*)
VAR_INPUT
	(* Variables *)
	bEnable								:BOOL;						(* Enable FB *)
	lrInSignal								:LREAL;						(* Input value to the block *)
	lrKp									:LREAL := 1;					(* Proportional gain of integrator *)
	tT1									:TIME := t#200ms;				(* Time constant  of integrator *)
	tTaskCycle							:TIME := t#2ms;				(* Cycle time *)
END_VAR
VAR_OUTPUT
	(* Variables *)
	lrOutSignal							:LREAL;						(* Output value the block state *)
END_VAR
VAR
	(* Variables *)
	bFirstTime							:BOOL;
	lrTimeRatio							:LREAL;

	lrLastSignal							:LREAL;						(* Last signal *)
END_VAR

IF NOT bEnable
THEN
	lrOutSignal := 0.0;
	bFirstTime := FALSE;
	RETURN;
END_IF


IF NOT bFirstTime
     OR tT1= t#0ms
     OR tT1 < (tTaskCycle + tTaskCycle)
THEN
	lrOutSignal := lrKp * lrInSignal;

	bFirstTime := TRUE;
ELSE
	lrTimeRatio := TIME_TO_LREAL(tTaskCycle) / TIME_TO_LREAL(tT1);

	lrOutSignal := (lrKp * lrInSignal * lrTimeRatio) + (lrLastSignal * (1 -  lrTimeRatio));
END_IF

lrLastSignal := lrOutSignal;

END_FUNCTION_BLOCK

// ---- POUs/Tc2 Objects/Engineering/Position offset/F_PosOffset.TcPOU
FUNCTION F_PosOffset : LREAL
(*

The function used to calculate position offset in range.

Constructor: 		Patryk Panylo
Company:		E. Riexinger GmbH
Date:			01.04.2015
Version:			1.00

Date:			Revision:		Who:				Comment
dd.mm.yyyy		x.xx			Initials			comment

*)
VAR_INPUT
	(* Input variables / Eingang Variablen *)
	bEnable							:BOOL;						(* Function enable *)
	lrCurrentPosHorizontal				:LREAL;						(* Current position of horizontal axis *)
	lrPosOffsetHorizontal				:LREAL;						(* Position offset of horizontal axis*)
	lrPosOffsetVertical					:LREAL;						(* Position offset of horizontal axis*)
	lrRangeOffset						:LREAL;						(* Range offset *)
END_VAR
VAR
	(* Variables *)

END_VAR

IF NOT bEnable
THEN
	F_PosOffset := 0.0;

	RETURN;
END_IF

IF  lrRangeOffset > 0.0
     AND lrCurrentPosHorizontal >= lrPosOffsetHorizontal - ABS(lrRangeOffset * 0.5)
     AND lrCurrentPosHorizontal <= lrPosOffsetHorizontal + ABS(lrRangeOffset * 0.5)
THEN
	F_PosOffset := lrPosOffsetVertical;
ELSE
	F_PosOffset := 0.0;
END_IF

END_FUNCTION

// ---- POUs/Tc2 Objects/Engineering/Position/F_ModuloDistance.TcPOU
FUNCTION F_ModuloDistance : DINT
(*
Function for calculate modulo distance.

Constructor: 	Patryk Panylo
Company:		E. Riexinger GmbH
Date:			20.01.2014
Version:		1.00

Date:			Revision:		Who:				Comment
dd.mm.yyyy		x.xx			Initials			comment

*)

VAR_INPUT
	dwCurrentValue			:DWORD;
	dwOldValue				:DWORD;
	dwModuloValue			:DWORD;
END_VAR
VAR
	dwPosDistance			:DWORD;

END_VAR


F_ModuloDistance := DWORD_TO_DINT(dwCurrentValue - dwOldValue);

IF dwModuloValue <> 0
THEN
	dwPosDistance := F_ModDW(dwCurrentValue - dwOldValue, dwModuloValue);
	
	F_ModuloDistance := DWORD_TO_DINT(dwPosDistance);
	
	IF dwPosDistance > (dwModuloValue / 2) 
	THEN
		F_ModuloDistance := -DWORD_TO_DINT(dwModuloValue - dwPosDistance);
	END_IF
	
END_IF

END_FUNCTION

// ---- POUs/Tc2 Objects/Mathematical/F_ModDW.TcPOU
FUNCTION F_ModDW : DWORD
(*
Modulo function for double word numbers (dividend mod divisor).

Constructor: 		Patryk Panylo
Company:		E. Riexinger GmbH
Date:			20.01.2014
Version:			1.00

Date:			Revision:		Who:				Comment
dd.mm.yyyy		x.xx			Initials			comment

*)
VAR_INPUT
	dwDividend						:DWORD;
	dwDivisor						:DWORD;
END_VAR
VAR
END_VAR


F_MODDW := dwDivisor;

IF dwDivisor <> 0 
THEN
	F_MODDW := dwDividend MOD dwDivisor;
END_IF;

END_FUNCTION

// ---- POUs/Tc2 Objects/Engineering/Trajectory model/FB_ExtContour.TcPOU
FUNCTION_BLOCK FB_ExtContour
(*

The function block used to generate move external contour.

Constructor: 		Patryk Panylo
Company:		E. Riexinger GmbH
Date:			01.04.2015
Version:			1.00

Date:			Revision:		Who:				Comment
dd.mm.yyyy		x.xx			Initials			comment

*)
VAR_INPUT
	(* Input variables / Eingang Variablen *)
	bEnable							:BOOL;						(* Function block enable *)
	bStart							:BOOL;
	bStop							:BOOL;
	etContourType					:ET_ContourType;				(* Contour type *)
	lrActPosZ						:LREAL;						(* Current position of axis z *)
	lrActAngle 						:LREAL; 						(* Current angle *)
	lrStartMaxPosZ					:LREAL;						(* Contour start maximal position of axis z *)
	lrEndMinPosZ					:LREAL;						(* Contour end minimal position of axis z *)
	lrSafetyDistance					:LREAL;						(* Safety distance *)
	lrTargetPosY						:LREAL;						(* Target position of axis y *)
END_VAR
VAR_OUTPUT
	(* Output variables / Ausgang Variablen *)
	lrNewPos						:LREAL;						(* New position [mm] *)
	bEnabled  						:BOOL;						(* Calculate positon is enabled *)
	lrActVelo							:LREAL;
	lrActPosN1						:LREAL;
END_VAR
VAR_IN_OUT
	lrSetPosY						:LREAL;						(* Set position of axis y *)
END_VAR
VAR
	(* Instances / Instanzen *)

	(* Enumerator  *)

	(* General flags / Allgemeine Variablen *)
	lrContourPos						:LREAL;
	bFirstTime						:BOOL;


END_VAR
VAR CONSTANT

END_VAR

IF NOT bEnable
THEN
	bEnabled := bStart;

	bFirstTime := FALSE;
	RETURN;
END_IF

IF NOT bFirstTime
THEN
	bEnabled := FALSE;

	bFirstTime := TRUE;
END_IF


IF bStop
THEN
	bEnabled := FALSE;

ELSIF bStart
THEN
	lrContourPos := F_CalcContour(
		etContourType := etContourType,
		lrActPos := lrActPosZ,
		lrActAngle := lrActAngle,
		(*lrActVelo := Axis.stNcToPlc.stCommandPositioning.dnActVelocity,*)
		lrVerticalOffset := 0.0,  (*37.0,*) (* Offset Sägeband Unterkante zu Störkontur BF-Kopf *)
		lrStartMaxPos := lrStartMaxPosZ,
		lrEndMinPos := lrEndMinPosZ,
		lrSafetyDistance := lrSafetyDistance,
		lrTableHeight := SEL(lrStartMaxPosZ>450, 700.0, 200.0), (* ab welcher Höhe Tischbreite aktiv ist *)
		lrTableWidth := 700.0, (* Tischbreite Auflage Rohr *)
		lrActVeloExt := lrActVelo
	);


	lrSetPosY := lrTargetPosY + lrContourPos;

	bEnabled := TRUE;

END_IF



lrActVelo := (*lrActVelo *0.9 + 0.1 *)(lrActPosZ - lrActPosN1);
lrActPosN1:= lrActPosZ;

END_FUNCTION_BLOCK

// ---- POUs/Tc2 Objects/Engineering/Trajectory model/F_CalcContour.TcPOU
FUNCTION F_CalcContour : LREAL
(*

The function used to calculate a contour of half circle dependent on angle of inclination axis and radius circle
Calculated position of axis is on output mapped.

Constructor: 		Patryk Panylo
Company:		E. Riexinger GmbH
Date:			01.04.2015
Version:			1.00

Date:			Revision:		Who:				Comment
dd.mm.yyyy		x.xx				Initials				comment
19.11.2015		1.01				ES					ET_ContourType_eEllipse
23.11.2015		1.02				ES					Square: also depending on angle(lrActAngle),
													lrVerticalOffset: guiding collision point is higher than act. position.

*)
VAR_INPUT
	(* Input variables / Eingang Variablen *)
	etContourType					:ET_ContourType;
	lrActPos							:LREAL;						(* Current position of axis *)
	lrActAngle						:LREAL;						(* Current angle, cutting angle *)
	(*lrActVelo							:LREAL;						(* Current speed of axis *)*)
	lrVerticalOffset					:LREAL;						(* vertical offset collision contour *)
	lrStartMaxPos						:LREAL;						(* Contour start maximal position *)
	lrEndMinPos						:LREAL;						(* Contour end minimal position  *)
	lrSafetyDistance					:LREAL;						(* Safety distance *)
	lrTableHeight						:LREAL;						(* Table height, if need guidings go to table width *)
	lrTableWidth						:LREAL;						(* table width *)
	lrActVeloExt						:LREAL;						(* Current velo of axis *)
END_VAR
VAR
	(* Variables *)
	lrActPosCache					:LREAL;						(* intern position of axis *)
	lrRadius							:LREAL;						(* Radius *)
	lrMiddlePos						:LREAL;						(* Middle position *)
	lrAlfa							:LREAL;						(* Angle of inclination *)
	lrDelta							:LREAL;						(* Distance z = f(x)*)
	lrCosAlfa							:LREAL;						(* Cosine of alfa *)
	lrAngleFactor						:LREAL;						(* Sawbow angle factor, ellipse *)
	lrStartMaxPosCache 				:LREAL;
	lrEndMinPosCache 				:LREAL;

END_VAR

lrStartMaxPosCache := lrStartMaxPos + ABS(lrSafetyDistance) + 50.0;
lrEndMinPosCache := lrEndMinPos - ABS(lrSafetyDistance) + 50.0;

lrActPosCache := lrActPos - lrVerticalOffset;

CASE etContourType OF

	ET_ContourType_eNone:
		F_CalcContour := lrActPosCache;

	ET_ContourType_eCircle, ET_ContourType_eEllipse:
		lrRadius := ABS(lrStartMaxPosCache - lrEndMinPos) / 2;
		lrMiddlePos := lrEndMinPosCache + lrRadius;										(* Middle position *)

		IF (lrActPosCache <= lrStartMaxPosCache)
		     AND (lrActPosCache >= lrEndMinPosCache)
		     AND lrRadius > 0.0
		THEN
			lrAlfa := ASIN(ABS(lrActPosCache - lrMiddlePos) /  lrRadius);				(* Angle of inclination *)
			lrCosAlfa := COS(lrAlfa);												(* Cosine of alfa *)
			lrDelta := lrCosAlfa * lrRadius;								(* Distance z = f(x)*)

			F_CalcContour := lrDelta;

		ELSE
			F_CalcContour := 0.0;
		END_IF

		IF lrActPos <= lrTableHeight
			OR lrActPos < lrMiddlePos
		THEN
			F_CalcContour := MAX(F_CalcContour, lrTableWidth / 2 + lrSafetyDistance);
		END_IF

		IF ((lrActVeloExt>0.0)
			AND (lrActPosCache < lrMiddlePos))
			OR ((lrActVeloExt=0.0)
			AND lrActPos < lrTableHeight)
		THEN
			F_CalcContour := MAX(lrRadius, lrTableWidth / 2 + lrSafetyDistance);
		END_IF

		IF etContourType = ET_ContourType_eEllipse
		THEN
			lrAngleFactor := 1 /  COS( MIN(ABS(lrActAngle), 89.9) / 180.0*PI);
			F_CalcContour := F_CalcContour * lrAngleFactor;
		END_IF

	ET_ContourType_eSquare:
		lrRadius := ABS(lrStartMaxPosCache - lrEndMinPos) / 2;
		lrMiddlePos := lrEndMinPosCache + lrRadius;										(* Middle position *)

		IF (lrActPosCache <= lrStartMaxPosCache)
		     AND (lrActPosCache >= lrEndMinPosCache)
		     AND lrRadius > 0.0
		THEN
			lrDelta := lrRadius;													(* Distance z = f(x)*)

			F_CalcContour := lrDelta;

		ELSE
			F_CalcContour := 0.0;
		END_IF

		IF lrActPos <= lrTableHeight
		THEN
			F_CalcContour := MAX(F_CalcContour, lrTableWidth / 2 + lrSafetyDistance / 2);
		END_IF

		lrAngleFactor := 1 /  COS( MIN(ABS(lrActAngle), 89.9) / 180.0*PI);
		F_CalcContour := F_CalcContour * lrAngleFactor;

ELSE
	F_CalcContour := 0.0;

END_CASE;

END_FUNCTION

// ---- POUs/Tc2 Objects/Engineering/Trajectory model/FB_ExtTraj.TcPOU
FUNCTION_BLOCK FB_ExtTraj
(*

The function block used to generate move external trajectory.

Constructor: 		Patryk Panylo
Company:		E. Riexinger GmbH
Date:			01.04.2015
Version:			1.00

Date:			Revision:		Who:				Comment
dd.mm.yyyy		x.xx			Initials			comment

*)
VAR_INPUT
	(* Input variables / Eingang Variablen *)
	bEnable							:BOOL;						(* Function block enable *)
	bStart							:BOOL;						(* Execute start an external trajectory with rising edge *)
	bStop							:BOOL;						(* Execute stop an external trajectory with rising edge *)
	lrStartPosHorizontal				:LREAL;						(* Start position of horizontal axis [mm] *)
	lrStartPosVertical					:LREAL;						(* Start position of vertical axis [mm] *)
	lrRadius							:LREAL;						(* Radius of circle [mm] *)
	unPosWindow					:UINT := 2;					(* Position window [mm] *)
	bTakeHorMovePara				:BOOL;						(* Take move parameters from 1- horizontal axis, 0 - vertical axis *)
END_VAR
VAR_OUTPUT
	(* Output variables / Ausgang Variablen *)
	lrNewPos						:LREAL;						(* New position [mm] *)
	lrNewVelo						:LREAL;						(* New velocity [mm/s] *)
	lrNewAcc						:LREAL;						(* New acceleration [mm/s^2] *)
	bEnabled  						:BOOL;						(* Calculate positon is enabled *)
	bDone							:BOOL;						(* Command done *)
	bBusy							:BOOL;						(* Command busy *)
	bError							:BOOL;						(* Command error  *)
	udnErrorNo						:UDINT;						(* Error number *)
	sErrorMsg						:STRING; 					(* Error message *)
END_VAR
VAR_IN_OUT
	AxisHorizontal					:AXIS_REF;					(* The AXIS_REF data type  is an interface between the PLC and the NC and contains axis information *)
	AxisVertical						:AXIS_REF;					(* The AXIS_REF data type  is an interface between the PLC and the NC and contains axis information *)
END_VAR
VAR
	(* Instances / Instanzen *)

	(* Enumerator  *)
	etCalcExtTrajState					:ET_CalcExtTrajState;								(* Current state *)

	(* General flags / Allgemeine Variablen *)
	lrExtStartPosHorizontal				:LREAL;
	lrExtStartPosVertical				:LREAL;
	lrExtRadius						:LREAL;

	bFirstTime						:BOOL;
END_VAR
VAR CONSTANT

END_VAR

IF NOT bEnable
THEN
	lrNewPos := SEL(bTakeHorMovePara, AxisVertical.NcToPlc.SetPos, AxisHorizontal.NcToPlc.SetPos);
	lrNewVelo := SEL(bTakeHorMovePara, AxisVertical.NcToPlc.SetVelo, AxisHorizontal.NcToPlc.SetVelo);
	lrNewAcc := SEL(bTakeHorMovePara, AxisVertical.NcToPlc.SetAcc, AxisHorizontal.NcToPlc.SetAcc);

	bDone := FALSE;					(* Command done *)
	bBusy := FALSE;					(* Command busy *)
	bError := FALSE;					(* Command error  *)
	udnErrorNo := 0;					(* Error number *)
	sErrorMsg := ''; 					(* Error message *)

	bEnabled := FALSE;

	bFirstTime := FALSE;
	RETURN;
END_IF

IF NOT bFirstTime
THEN
	bEnabled := FALSE;

	etCalcExtTrajState := ET_CalcExtTrajState_eWaitExecute;

	bFirstTime := TRUE;
END_IF

CASE etCalcExtTrajState
OF
	ET_CalcExtTrajState_eWaitExecute:
		IF bStop
		THEN
			bEnabled := FALSE;

			bDone := FALSE;						(* Command done *)
			bBusy := TRUE;						(* Command busy *)
			bError := FALSE;						(* Command error  *)
			udnErrorNo := 0;						(* Error number *)
			sErrorMsg := ''; 						(* Error message *)

			etCalcExtTrajState := ET_CalcExtTrajState_eDone;

		ELSIF bStart
		THEN
			bDone := FALSE;						(* Command done *)
			bBusy := TRUE;						(* Command busy *)
			bError := FALSE;						(* Command error  *)
			udnErrorNo := 0;						(* Error number *)
			sErrorMsg := ''; 						(* Error message *)

			etCalcExtTrajState := ET_CalcExtTrajState_eCalcTrajPos;

		END_IF

	ET_CalcExtTrajState_eCalcTrajPos:
		bEnabled := TRUE;

		lrExtStartPosHorizontal := lrStartPosHorizontal;
		lrExtStartPosVertical := lrStartPosVertical;
		lrExtRadius := lrRadius;

		etCalcExtTrajState := ET_CalcExtTrajState_eDone;

	ET_CalcExtTrajState_eError:
		bBusy := FALSE;						(* Command busy *)
		bError := TRUE;						(* Command error  *)

		etCalcExtTrajState := ET_CalcExtTrajState_eNoExecute;

	ET_CalcExtTrajState_eDone:
		bDone := TRUE;						(* Command done *)
		bBusy := FALSE;						(* Command busy *)

		etCalcExtTrajState := ET_CalcExtTrajState_eNoExecute;

	ET_CalcExtTrajState_eNoExecute:
		IF NOT bStart
		     AND NOT bStop
		THEN
			(* Reset outputs *)
			bDone := FALSE;						(* Command done *)
			bBusy := FALSE;						(* Command busy *)
			bError := FALSE;						(* Command error  *)

			etCalcExtTrajState := ET_CalcExtTrajState_eWaitExecute;
		END_IF
END_CASE

(* The function is used to calculate a trajectory of vertical position. *)
IF bEnabled
THEN
	lrNewPos := F_CalcTrajPos(
		lrStartPosHorizontal := lrExtStartPosHorizontal,
		lrStartPosVertical := lrExtStartPosVertical,
		lrCurrentPosHorizontal := AxisHorizontal.NcToPlc.SetPos,
		lrCurrentPosVertical := AxisVertical.NcToPlc.SetPos,
		lrRadius := lrExtRadius
	);

	lrNewVelo := AxisHorizontal.NcToPlc.SetVelo;
	lrNewAcc := AxisHorizontal.NcToPlc.SetAcc;

	(* ABS(lrNewPos - AxisVertical.NcToPlc.SetPos) > UINT_TO_LREAL(unPosWindow)
	THEN
		bError := TRUE;								(* Command error  *)
		udnErrorNo :=  1;								(* Error number *)
		sErrorMsg := ''; 								(* Error message *)
	END_IF*)
ELSE
	lrNewPos := SEL(bTakeHorMovePara, AxisVertical.NcToPlc.SetPos, AxisHorizontal.NcToPlc.SetPos);
	lrNewVelo := SEL(bTakeHorMovePara, AxisVertical.NcToPlc.SetVelo, AxisHorizontal.NcToPlc.SetVelo);
	lrNewAcc := SEL(bTakeHorMovePara, AxisVertical.NcToPlc.SetAcc, AxisHorizontal.NcToPlc.SetAcc);

	bError := FALSE;								(* Command error  *)
	udnErrorNo :=  0;								(* Error number *)
	sErrorMsg := ''; 								(* Error message *)
END_IF

END_FUNCTION_BLOCK

// ---- POUs/Tc2 Objects/Engineering/Trajectory model/F_CalcTrajPos.TcPOU
FUNCTION F_CalcTrajPos : LREAL
(*

The function used to calculate a trajectory of half circle dependent on angle of inclination axis and radius circle
Calculated position of axis is on output mapped.

Constructor: 		Patryk Panylo
Company:		E. Riexinger GmbH
Date:			01.04.2015
Version:			1.00

Date:			Revision:		Who:				Comment
dd.mm.yyyy		x.xx			Initials			comment

*)
VAR_INPUT
	(* Input variables / Eingang Variablen *)
	lrStartPosHorizontal				:LREAL;						(* Start position of horizontal axis *)
	lrStartPosVertical					:LREAL;						(* Start position of vertical axis *)
	lrCurrentPosHorizontal				:LREAL;						(* Current position of horizontal axis *)
	lrCurrentPosVertical				:LREAL;						(* Current position of vertical axis *)
	lrRadius							:LREAL;						(* Radius of circle *)
END_VAR
VAR
	(* Variables *)
	lrAlfa							:LREAL;						(* Angle of inclination *)
	lrDelta							:LREAL;						(* Distance z = f(x)*)
	lrCosAlfa							:LREAL;						(* Cosine of alfa *)
END_VAR

IF lrRadius > 0.0
THEN
	IF ABS(lrCurrentPosHorizontal - lrStartPosHorizontal) / lrRadius <= 1.0
	THEN
		lrAlfa := ASIN(ABS(lrCurrentPosHorizontal - lrStartPosHorizontal) / lrRadius);					(* Angle of inclination *)
		lrCosAlfa := COS(lrAlfa);																(* Cosine of alfa *)
		lrDelta := lrRadius - (lrCosAlfa * lrRadius);											(* Distance z = f(x)*)

		F_CalcTrajPos := lrCurrentPosVertical - lrDelta;
	ELSE
		F_CalcTrajPos := lrCurrentPosVertical;
	END_IF
ELSE
	F_CalcTrajPos := lrCurrentPosVertical;
END_IF

END_FUNCTION

// ---- POUs/Tc2 Objects/ExternalHardware/Gefran/FB_GFX4IRCtrlZone.TcPOU
FUNCTION_BLOCK FB_GFX4IRCtrlZone
(*

The function block used to control Gerfan GFX4IR zone.

Constructor: 		Patryk Panylo
Company:		E. Riexinger GmbH
Date:			12.07.2016
Version:			1.00

Date:			Revision:		Who:				Comment
13.12.2017		1.01				PPA					Control with temperatur feedback

*)
VAR_INPUT
	(* Input variables / Eingang Variablen *)
	bEnable							:BOOL;						(* Function block enable *)
	bReset							:BOOL;						(* Controller reset *)
	bHandStart						:BOOL;						(* Execute start an external trajectory with rising edge *)
	bHandStop						:BOOL;						(* Execute stop an external trajectory with rising edge *)
	bAutoStart						:BOOL;						(* Execute start an external trajectory with rising edge *)
	bAutoStop						:BOOL;						(* Execute stop an external trajectory with rising edge *)
	bStartRelease					:BOOL;						(* Start release *)
	bCtrlInterrupt						:BOOL;						(* Control interrupt *)
	lrSetpoint						:LREAL;						(* Setpoint *)
	bCtrlManAuto						:BOOL;						(* Auto := FALSE, Man := TRUE *)
	bEnAutoCtrlOff					:BOOL := TRUE;				(* Auto off enable*)
	tControllerOff						:TIME := t#90s;				(* Time to switch controller off *)
	tControllerOn						:TIME := t#90s;				(* Time to switch controller on *)
	lrTempMin						:LREAL;						(* Minimal temperature *)
	lrTempMax						:LREAL;						(* Maximal temperature *)
	lrTempLimitMin					:LREAL;						(* Minimal temperature limit *)
	lrTempLimitMax					:LREAL;						(* Maximal temperature limit *)
END_VAR
VAR_OUTPUT
	(* Output variables / Ausgang Variablen *)
	unCurrentValue					:UINT;						(* Current value *)
	bEnabled  						:BOOL;						(* Zone enabled *)
	bDamaged						:BOOL;						(* Zone damaged *)
	bDone							:BOOL;						(* Command done *)
	bBusy							:BOOL;						(* Command busy *)
	bError							:BOOL;						(* Command error  *)
	udnErrorNo						:UDINT;						(* Error number *)
	sErrorMsg						:STRING; 					(* Error message *)
END_VAR
VAR_IN_OUT
	(* Input Output variables / Ausgang Variablen *)
	CtrlGFX4IRTOPLC					:ST_GFX4IRTOPLC;			(* The ST_GFX4IRTOPLC data type  is an interface between the PLC and the GFX4IR and contains controller information *)
	CtrlPLCTOGFX4IR					:ST_PLCTOGFX4IR;			(* The ST_PLCTOGFX4IR data type  is an interface between the PLC and the GFX4IR and contains controller information *)
END_VAR
VAR
	(* Enummerations *)
	etGFX4IRStates					:ET_GFX4IR := ET_GFX4IRState_eWaitExecute;			(* Current state *)

	(* Variables *)
	nWatchdog						:INT;
	bControllerOn						:BOOL;

	bFirstTime						:BOOL;

	(* References *)

	(* Interfaces *)

	(* Instances *)
	fbControllerOff					:FB_SignalHandlingDelay;
	fbControllerOn					:FB_SignalHandlingDelay;
	fbScalingSP						:FB_Scaling;

	rtAutoStart						:R_TRIG;
	rtAutoStop						:R_TRIG;
	rtHandStart						:R_TRIG;
	rtHandStop						:R_TRIG;
END_VAR
VAR CONSTANT

END_VAR


IF NOT bFirstTime
THEN
	bControllerOn := TRUE;

	nWatchdog := 0;
	bDone := FALSE;						(* Command done *)
	bBusy := FALSE;						(* Command busy *)
	bError := FALSE;						(* Command error  *)

	etGFX4IRStates := ET_GFX4IRState_eWaitExecute;

	bFirstTime := TRUE;
END_IF

(* Scaling set point *)
fbScalingSP(
	bEnable := TRUE,
	lrInput := lrSetpoint,
	lrXLowLimit := lrTempMin,
	lrXUpperLimit := lrTempMax,
	lrYLowLimit := lrTempLimitMin,
	lrYUpperLimit := lrTempLimitMax,
	usiPrecision := 2
);

CtrlPLCTOGFX4IR.wControllerStatus.4 := bCtrlManAuto;			(* Auto := FALSE, Man := TRUE *)

IF bCtrlManAuto										(* Auto := FALSE, Man := TRUE *)
THEN
	bEnabled := CtrlGFX4IRTOPLC.nOutputPower > 0
			       AND (CtrlGFX4IRTOPLC.nOutputPower = LREAL_TO_INT(lrSetpoint  * 10.0));
			       (*AND CtrlGFX4IRTOPLC.wControllerStatus.5					(* Ctrl enabled  *)
			          AND NOT CtrlGFX4IRTOPLC.wControllerStatus.0;			(* Alarm  *)*)
ELSE
	bEnabled := CtrlGFX4IRTOPLC.nOutputPower > 0;
			       (*AND (CtrlGFX4IRTOPLC.nProcessVariable >= LREAL_TO_INT(fbScalingSP.lrOutputPV));*)
			       (*AND CtrlGFX4IRTOPLC.wControllerStatus.5					(* Ctrl enabled  *)
			          AND NOT CtrlGFX4IRTOPLC.wControllerStatus.0;			(* Alarm  *)*)
END_IF

bDamaged := CtrlGFX4IRTOPLC.wControllerStatus.12;
unCurrentValue := CtrlGFX4IRTOPLC.nOutputPower / 10;

fbControllerOff(
	bEnable := TRUE,
	bIn := bEnAutoCtrlOff
		  AND bEnabled,
	tDelay := tControllerOff
);

fbControllerOn(
	bEnable := TRUE,
	bIn := NOT bEnabled					(* Ctrl disabled *)
		  AND NOT bControllerOn,
	tDelay := tControllerOn
);

(*
IF bHandStop
    OR bCtrlInterrupt
THEN
	CtrlPLCTOGFX4IR.wControllerStatus.3 := TRUE;			(* Ctrl ON = FALSE, OFF = TRUE *)
	CtrlPLCTOGFX4IR.nLocalSetPoint := 0;
	CtrlPLCTOGFX4IR.nManualOutput := 0;
ELSIF bHandStart
THEN
	CtrlPLCTOGFX4IR.wControllerStatus.3 := FALSE;			(* Ctrl ON = FALSE, OFF = TRUE *)
	CtrlPLCTOGFX4IR.nManualOutput := LREAL_TO_INT(lrSetpoint  * 10);
END_IF

RETURN;
*)

IF bCtrlInterrupt
     OR fbControllerOff.bOut
THEN
	bControllerOn := FALSE;

	CtrlPLCTOGFX4IR.wControllerStatus.3 := TRUE;			(* Ctrl ON = FALSE, OFF = TRUE *)
	CtrlPLCTOGFX4IR.nLocalSetPoint := 0;
	CtrlPLCTOGFX4IR.nManualOutput := 0;

	nWatchdog := 0;
	bDone := FALSE;						(* Command done *)
	bBusy := FALSE;						(* Command busy *)
	bError := FALSE;						(* Command error  *)

	etGFX4IRStates := ET_GFX4IRState_eWaitExecute;

ELSIF fbControllerOn.bOut
THEN
	bControllerOn := TRUE;
END_IF

IF bReset
     AND bError
THEN
	(* Reset outputs *)
	nWatchdog := 0;
	bDone := FALSE;						(* Command done *)
	bBusy := FALSE;						(* Command busy *)
	bError := FALSE;						(* Command error  *)

	etGFX4IRStates := ET_GFX4IRState_eWaitExecute;
ELSE
	(*IF bEnable
	     AND CtrlGFX4IRTOPLC.wControllerStatus.8					(* Ctrl error *)
	THEN
		bError := TRUE;									(* Command error  *)

		etGFX4IRStates := ET_GFX4IRState_eError;             		(* Next step *)
	END_IF*);
END_IF

rtHandStart(CLK := bHandStart);
rtHandStop(CLK := bHandStop);
rtAutoStart(CLK := bAutoStart AND bStartRelease AND bControllerOn);
rtAutoStop(CLK := bAutoStop);

IF rtHandStart.Q OR rtHandStop.Q
     OR rtAutoStart.Q OR rtAutoStop.Q
THEN
	nWatchdog := 0;
	bDone := FALSE;						(* Command done *)
	bBusy := FALSE;						(* Command busy *)
	bError := FALSE;						(* Command error  *)

	etGFX4IRStates := ET_GFX4IRState_eWaitExecute;
END_IF

CASE etGFX4IRStates
OF
	ET_GFX4IRState_eWaitExecute:
		IF NOT bEnable
		THEN
			bDone := TRUE;						(* Command done *)
			bBusy := TRUE;						(* Command busy *)
			bError := FALSE;						(* Command error  *)
			bEnabled  := bAutoStart AND NOT bAutoStop; 				(* Controller enabled *)

			etGFX4IRStates := ET_GFX4IRState_eWaitExecute;

		ELSIF NOT bCtrlInterrupt
			    AND NOT fbControllerOff.bOut
		THEN
			IF bAutoStop
			     OR bHandStop
			THEN
				nWatchdog := 0;

				bDone := FALSE;						(* Command done *)
				bBusy := TRUE;						(* Command busy *)
				bError := FALSE;						(* Command error  *)
				udnErrorNo := 0;						(* Error number *)
				sErrorMsg := ''; 						(* Error message *)

				etGFX4IRStates := ET_GFX4IRState_eCtrlOff;

			ELSIF rtAutoStart.Q
				    OR (rtHandStart.Q
					    AND bStartRelease
					    AND bControllerOn)
			THEN
				nWatchdog := 0;

				bDone := FALSE;						(* Command done *)
				bBusy := TRUE;						(* Command busy *)
				bError := FALSE;						(* Command error  *)
				udnErrorNo := 0;						(* Error number *)
				sErrorMsg := ''; 						(* Error message *)

				etGFX4IRStates := ET_GFX4IRState_eCtrlOn;

			END_IF
		END_IF

	ET_GFX4IRState_eCtrlOn:
		nWatchdog := nWatchdog + 1;

		CtrlPLCTOGFX4IR.wControllerStatus.3 := FALSE;			(* Ctrl ON = FALSE, OFF = TRUE *)

		IF bCtrlManAuto										(* Auto := FALSE, Man := TRUE *)
		THEN
			CtrlPLCTOGFX4IR.nManualOutput := LREAL_TO_UINT(lrSetpoint  * 10.0);
		ELSE
			CtrlPLCTOGFX4IR.nLocalSetPoint := LREAL_TO_INT(fbScalingSP.lrOutputPV);
		END_IF

		IF bEnabled											(* Ctrl enabled *)
		THEN
			nWatchdog := 0;
			etGFX4IRStates := ET_GFX4IRState_eDone;

		ELSIF nWatchdog > 5000
		THEN
			CtrlPLCTOGFX4IR.wControllerStatus.3 := TRUE;			(* Ctrl ON = FALSE, OFF = TRUE *)

			etGFX4IRStates := ET_GFX4IRState_eError;            		 (* Next step *)
		END_IF

	ET_GFX4IRState_eCtrlOff:
		nWatchdog := nWatchdog + 1;

		CtrlPLCTOGFX4IR.wControllerStatus.3 := TRUE;			(* Ctrl ON = FALSE, OFF = TRUE *)
		CtrlPLCTOGFX4IR.nLocalSetPoint := 0;
		CtrlPLCTOGFX4IR.nManualOutput := 0;

		IF NOT bEnabled
		THEN
			nWatchdog := 0;
			etGFX4IRStates := ET_GFX4IRState_eDone;

		ELSIF nWatchdog > 1000
		THEN
			CtrlPLCTOGFX4IR.wControllerStatus.3 := TRUE;			(* Ctrl ON = FALSE, OFF = TRUE *)
			CtrlPLCTOGFX4IR.nLocalSetPoint := 0;
			CtrlPLCTOGFX4IR.nManualOutput := 0;
			etGFX4IRStates := ET_GFX4IRState_eError;             		(* Next step *)
		END_IF

	ET_GFX4IRState_eDone:
		nWatchdog := 0;
		bDone := TRUE;						(* Command done *)
		bBusy := FALSE;						(* Command busy *)

		etGFX4IRStates := ET_GFX4IRState_eNoExecute;

	ET_GFX4IRState_eError:
		nWatchdog := 0;
		bBusy := FALSE;						(* Command busy *)
		bError := TRUE;						(* Command error  *)

		CtrlPLCTOGFX4IR.wControllerStatus.3 := TRUE;			(* Ctrl ON = FALSE, OFF = TRUE *)
		CtrlPLCTOGFX4IR.nLocalSetPoint := 0;
		CtrlPLCTOGFX4IR.nManualOutput := 0;

		etGFX4IRStates := ET_GFX4IRState_eNoExecute;

	ET_GFX4IRState_eNoExecute:
		IF NOT bHandStart
		     AND NOT bHandStop
		     AND NOT bAutoStart
		     AND NOT bAutoStop
		THEN
			(* Reset outputs *)
			nWatchdog := 0;
			bDone := FALSE;						(* Command done *)
			bBusy := FALSE;						(* Command busy *)
			bError := FALSE;						(* Command error  *)

			etGFX4IRStates := ET_GFX4IRState_eWaitExecute;
		END_IF
END_CASE

END_FUNCTION_BLOCK

// ---- POUs/Tc2 Objects/ExternalHardware/Gefran/FB_GFX4IRZones.TcPOU
FUNCTION_BLOCK FB_GFX4IRZones
(*

The function block used to control Gerfan GFX4IR Zones.

Constructor: 		Patryk Panylo
Company:		E. Riexinger GmbH
Date:			12.07.2016
Version:			1.00

Date:			Revision:		Who:				Comment
25.09.2017		1.01				PPA					Change check zone damaged

*)
VAR_INPUT
	(* Input variables / Eingang Variablen *)
	bEnable							:BOOL;													(* Function block enable *)
	arbZoneEn						:ARRAY[1..nZONES_MAX_NO] OF BOOL;						(* Zone enable *)
	bReset							:BOOL;													(* Reset *)
	arbHandStart						:ARRAY[1..nZONES_MAX_NO] OF BOOL;						(* Execute start GFX4IR controller with rising edge *)
	arbHandStop						:ARRAY[1..nZONES_MAX_NO] OF BOOL;						(* Execute stop GFX4IR controller with rising edge *)
	bAutoStart						:BOOL;													(* Execute start GFX4IR controller with rising edge *)
	bAutoStop						:BOOL;													(* Execute stop GFX4IR controller with rising edge *)
	bStartRelease					:BOOL;													(* Start release *)
	bCtrlInterrupt						:BOOL;													(* Control interrupt *)
	arlrSetpoint						:ARRAY[1..nZONES_MAX_NO] OF LREAL;					(* Setpoint *)
	bCtrlManAuto						:BOOL;													(* Auto := FALSE, Man := TRUE *)
	bEnAutoCtrlOff					:BOOL := TRUE;											(* Auto controller off enable*)
	bEnOneByOneOn					:BOOL := FALSE;											(* One by one switch on *)
	tDelayZoneOn					:TIME := t#100ms;											(* Delay time of zone one by one to switch on *)
	tControllerOff						:TIME := t#90s;											(* Time to switch controller off *)
	tControllerOn						:TIME := t#90s;											(* Time to switch controller on *)
	lrTempMin						:LREAL;													(* Minimal temperature *)
	lrTempMax						:LREAL;													(* Maximal temperature *)
	lrTempLimitMin					:LREAL;													(* Minimal temperature limit *)
	lrTempLimitMax					:LREAL;													(* Maximal temperature limit *)
END_VAR
VAR_OUTPUT
	(* Output variables / Ausgang Variablen *)
	arunCurrentValue					:ARRAY[1..nZONES_MAX_NO] OF UINT;						(* Current value *)
	bEnabled  						:BOOL;													(* Zone enabled *)
	bEnabledDelay					:BOOL;													(* Zone enabled delay *)
	arbZoneDamaged				:ARRAY[1..nZONES_MAX_NO] OF BOOL;
	bDone							:BOOL;						(* Command done *)
	bError							:BOOL;						(* Command error  *)
	udnErrorNo						:UDINT;						(* Error number *)
END_VAR
VAR_IN_OUT
	(* Input Output variables / Ausgang Variablen *)
	GFX4IR							:ST_GFX4IR_REF;				(* The ST_GFX4IR_REF data type  is an interface between the PLC and the GFX4IR and contains controller information *)
END_VAR
VAR
	(* Enummerations *)

	(* Variables *)
	nIdx								:INT;
	tEnabledDelay					:TIME := t#1s;					(* Enabled delay time *)


	bFirstTime						:BOOL;

	(* References *)

	(* Interfaces *)

	(* Instances *)
	arfbGFX4IRCtrlZone				:ARRAY[1..nZONES_MAX_NO] OF FB_GFX4IRCtrlZone;
	tonEnabledDelay					:TON;						(* Delay controller enabled status *)
	tonDelayZoneOn					:ARRAY[1..nZONES_MAX_NO] OF TON;						(* Delay zone one by one to switch on *)

END_VAR


IF NOT bEnable
THEN
	bDone := FALSE;					(* Command done *)
	bError := FALSE;					(* Command error  *)

	FOR nIdx := 1 TO nZONES_MAX_NO
	DO
		arfbGFX4IRCtrlZone[nIdx](
			bEnable := TRUE,
			bAutoStart := bAutoStart,
			bAutoStop := bAutoStop,
			bCtrlInterrupt := bCtrlInterrupt,
			lrTempMin := lrTempMin,
			lrTempMax := lrTempMax,
			lrTempLimitMin := lrTempLimitMin,
			lrTempLimitMax := lrTempLimitMax,
			CtrlGFX4IRTOPLC := GFX4IR.Gfx4IRToPlc[nIdx],
			CtrlPLCTOGFX4IR := GFX4IR.PlcToGfx4IR[nIdx],
			unCurrentValue => arunCurrentValue[nIdx]
		 );
	END_FOR

	bEnabled := FALSE;
	bEnabledDelay := FALSE;

	bFirstTime := FALSE;
	RETURN;
END_IF

IF NOT bFirstTime
THEN
	bDone := FALSE;					(* Command done *)
	bError := FALSE;					(* Command error  *)

	bEnabled := FALSE;
	bEnabledDelay := FALSE;

	bFirstTime := TRUE;
END_IF

bEnabled := TRUE;
bDone := TRUE;
bError := FALSE;

FOR nIdx := 1 TO nZONES_MAX_NO
DO
	(*
	IF bAutoStart
	THEN
		IF bEnOneByOneOn
		     AND tDelayZoneOn > t#0ms
		     AND nIdx > 1
		     AND NOT arfbGFX4IRController[nIdx].bEnabled
		THEN
			tonDelayZoneOn[nIdx](
				IN := arfbGFX4IRController[nIdx - 1].bEnabled,
				PT := tDelayZoneOn
			);
	
			IF tonDelayZoneOn[nIdx].Q
			THEN
				arfbGFX4IRController[nIdx].bStartRelease := bStartRelease;
			ELSE
				arfbGFX4IRController[nIdx].bStartRelease := FALSE;;
			END_IF
		ELSE
			tonDelayZoneOn[nIdx](IN := FALSE);
			arfbGFX4IRController[nIdx].bStartRelease := bStartRelease;
		END_IF
	ELSE
		tonDelayZoneOn[nIdx](IN := FALSE);
		arfbGFX4IRController[nIdx].bStartRelease := bStartRelease;
	END_IF
	*)

	arfbGFX4IRCtrlZone[nIdx].bStartRelease := bStartRelease;

	arfbGFX4IRCtrlZone[nIdx](
		bEnable := arbZoneEn[nIdx],
		bReset := bReset,
		bHandStart := arbHandStart[nIdx],
		bHandStop := arbHandStop[nIdx],
		bAutoStart := bAutoStart,
		bAutoStop := bAutoStop,
		bCtrlInterrupt := bCtrlInterrupt,
		lrSetpoint := arlrSetpoint[nIdx],
		bCtrlManAuto := bCtrlManAuto,
		bEnAutoCtrlOff := bEnAutoCtrlOff,
		tControllerOff := tControllerOff,
		tControllerOn := tControllerOn,
		lrTempMin := lrTempMin,
		lrTempMax := lrTempMax,
		lrTempLimitMin := lrTempLimitMin,
		lrTempLimitMax := lrTempLimitMax,
		CtrlGFX4IRTOPLC := GFX4IR.Gfx4IRToPlc[nIdx],
		CtrlPLCTOGFX4IR := GFX4IR.PlcToGfx4IR[nIdx],
		unCurrentValue => arunCurrentValue[nIdx],
		bDamaged => arbZoneDamaged[nIdx]
	 );

	bEnabled := bEnabled AND arfbGFX4IRCtrlZone[nIdx].bEnabled;
	bDone := bDone AND arfbGFX4IRCtrlZone[nIdx].bDone;
	bError := bError OR arfbGFX4IRCtrlZone[nIdx].bError;

END_FOR

tonEnabledDelay(
	IN := bEnabled,
	PT := tEnabledDelay,
	Q => bEnabledDelay
);

END_FUNCTION_BLOCK

// ---- POUs/Tc2 Objects/ExternalHardware/Gefran/FB_GFX4IR_REF.TcPOU
FUNCTION_BLOCK FB_GFX4IR_REF
VAR_INPUT
	Gfx4IRToPlc			AT %I*:ARRAY[1..4] OF ST_GFX4IRTOPLC;
END_VAR
VAR_OUTPUT
	PlcToGfx4IR			AT %Q*:ARRAY[1..4] OF ST_PLCTOGFX4IR;
END_VAR
VAR
END_VAR

;

END_FUNCTION_BLOCK

// ---- POUs/Tc2 Objects/ExternalHardware/Gefran/F_ChkAllZonesNotEnabled.TcPOU
FUNCTION F_ChkAllZonesNotEnabled : BOOL
(*

The function used to detect if all controller are enabled.

Constructor: 		Patryk Panylo
Company:		E. Riexinger GmbH
Date:			23.04.2015
Version:			1.00

Date:			Revision:		Who:				Comment
dd.mm.yyyy		x.xx			Initials			comment

*)
VAR_INPUT
	(* Input variables / Eingang Variablen *)
	bEnable						:BOOL;						(* Signal FB enable *)
	GFX4IR1						:ST_GFX4IR_REF;				(* The ST_GFX4IRTOPLC data type  is an interface between the PLC and the GFX4IR and contains controller information *)
	GFX4IR2						:ST_GFX4IR_REF;				(* The ST_GFX4IRTOPLC data type  is an interface between the PLC and the GFX4IR and contains controller information *)
	GFX4IR3						:ST_GFX4IR_REF;				(* The ST_GFX4IRTOPLC data type  is an interface between the PLC and the GFX4IR and contains controller information *)
	GFX4IR4						:ST_GFX4IR_REF;				(* The ST_GFX4IRTOPLC data type  is an interface between the PLC and the GFX4IR and contains controller information *)
END_VAR
VAR
	(* Enummerations *)

	(* Variables *)

	(* References *)

	(* Interfaces *)

	(* Instances *)

END_VAR


IF NOT bEnable							(* Signal FB enable *)
THEN
	F_ChkAllZonesNotEnabled := FALSE;

	RETURN;
END_IF

F_ChkAllZonesNotEnabled := GFX4IR1.Gfx4IRToPlc[1].nProcessVariable = 0
						   AND GFX4IR1.Gfx4IRToPlc[2].nProcessVariable = 0
						   AND GFX4IR1.Gfx4IRToPlc[3].nProcessVariable = 0
						   AND GFX4IR1.Gfx4IRToPlc[4].nProcessVariable = 0
						   AND GFX4IR2.Gfx4IRToPlc[1].nProcessVariable = 0
						   AND GFX4IR2.Gfx4IRToPlc[2].nProcessVariable = 0
						   AND GFX4IR2.Gfx4IRToPlc[3].nProcessVariable = 0
						   AND GFX4IR2.Gfx4IRToPlc[4].nProcessVariable = 0
						   AND GFX4IR3.Gfx4IRToPlc[1].nProcessVariable = 0
						   AND GFX4IR3.Gfx4IRToPlc[2].nProcessVariable = 0
						   AND GFX4IR3.Gfx4IRToPlc[3].nProcessVariable = 0
						   AND GFX4IR3.Gfx4IRToPlc[4].nProcessVariable = 0
						   AND GFX4IR4.Gfx4IRToPlc[1].nProcessVariable = 0
						   AND GFX4IR4.Gfx4IRToPlc[2].nProcessVariable = 0
						   AND GFX4IR4.Gfx4IRToPlc[3].nProcessVariable = 0
						   AND GFX4IR4.Gfx4IRToPlc[4].nProcessVariable = 0;

END_FUNCTION

// ---- POUs/Tc2 Objects/ExternalHardware/KUKA/FB_KUKA_Enable.TcPOU
FUNCTION_BLOCK FB_KUKA_Enable
(*

The function block used to move enable for an kuka

Constructor: 		Patryk Panylo
Company:		E. Riexinger GmbH
Date:			18.11.2016
Version:			1.00

Date:			Revision:		Who:				Comment

*)
VAR_INPUT
	(* Input variables / Eingang Variablen *)
	bEnable						:BOOL;			(* Signal FB enable *)
	bAutoHand					:BOOL;			(* Auto := TRUE, Hand := FALSE *)
	bNoEStop					:BOOL;			(* No ermergency Stop / Keine Notaus *)
	bMoveOn					:BOOL;			(* Enable the move enable *)
END_VAR
VAR_OUTPUT
	(* Output variables / Ausgang Variablen *)
	bMoveEnabled				:BOOL;			(* MoveEnabled = TRUE indicates that the kuka  drivers is ready for operation. *)
	bError						:BOOL;			(* Error *)
	udnErrorNo					:UDINT;			(* Error number *)
	sErrorMsg					:STRING; 		(* Error message *)
END_VAR
VAR_IN_OUT
	(* Input Output variables / Ausgang Variablen *)
	Kuka							:ST_KUKA_REF;
END_VAR
VAR
	(* Enummerations *)

	(* Variables *)
	tMoveEnabledDelay 					:TIME := t#300ms;

	(* References *)

	(* Interfaces *)

	(* Instances *)
	tonMoveEnabledDelay					:TON;
END_VAR


IF NOT bEnable
THEN
	Kuka.PlcToKuka.bMoveEnable := FALSE;                   		 (* Disable *)
	tonMoveEnabledDelay(IN := FALSE,
				    		 PT := tMoveEnabledDelay);
ELSE

	IF NOT bNoEStop
	THEN
		Kuka.PlcToKuka.bMoveEnable := FALSE;                   		 (* Disable *)

	ELSE
		IF bAutoHand			(* Auto *)
		THEN
			IF (bMoveOn
			      OR (NOT bMoveOn
				     AND Kuka.KukaToPlc.bInWorkArea))
			     AND Kuka.KukaToPlc.bIOActConf
			     AND Kuka.KukaToPlc.bExt
			THEN
				Kuka.PlcToKuka.bMoveEnable := TRUE;                   		 (* Enable *)
			ELSE
				Kuka.PlcToKuka.bMoveEnable := FALSE;                   		 (* Enable *)
			END_IF
		ELSE				(* Manual *)
			IF Kuka.KukaToPlc.bT1
			     OR Kuka.KukaToPlc.bT2
			     OR Kuka.KukaToPlc.bAut
			THEN
				Kuka.PlcToKuka.bMoveEnable := TRUE;                   		 (* Enable *)
			ELSE
				Kuka.PlcToKuka.bMoveEnable := FALSE;                   		 (* Enable *)
			END_IF
		END_IF
	END_IF;

END_IF;

tonMoveEnabledDelay(IN := Kuka.PlcToKuka.bMoveEnable,				(* Move enabled *)
			   		PT := tMoveEnabledDelay);
bMoveEnabled := tonMoveEnabledDelay.Q;

END_FUNCTION_BLOCK

// ---- POUs/Tc2 Objects/ExternalHardware/KUKA/FB_KUKA_Power.TcPOU
FUNCTION_BLOCK FB_KUKA_Power
(*

The function block used to enable drives for an kuka

Constructor: 		Patryk Panylo
Company:		E. Riexinger GmbH
Date:			18.11.2016
Version:			1.00

Date:			Revision:		Who:				Comment

*)
VAR_INPUT
	(* Input variables / Eingang Variablen *)
	bEnable						:BOOL;			(* Signal FB enable *)
	bNoEStop					:BOOL;			(* No ermergency Stop / Keine Notaus *)
	bDrivesOn					:BOOL;			(* Enable the drives *)
	lrOverride					:LREAL;			(* Velocity override in % for all motion commands. (0 <= Override <= 100.0) *)
END_VAR
VAR_OUTPUT
	(* Output variables / Ausgang Variablen *)
	bStatus						:BOOL;			(* Status = TRUE indicates that the axis is ready for operation. *)
	bError						:BOOL;			(* Error *)
	udnErrorNo					:UDINT;			(* Error number *)
	sErrorMsg					:STRING; 		(* Error message *)
END_VAR
VAR_IN_OUT
	(* Input Output variables / Ausgang Variablen *)
	Kuka						:ST_KUKA_REF;
END_VAR
VAR
	(* Enummerations *)

	(* Variables *)
	tStatusDelay 					:TIME := t#300ms;

	(* References *)

	(* Interfaces *)

	(* Instances *)
	tonStatusDelay				:TON;
END_VAR


IF NOT bEnable
THEN
	Kuka.PlcToKuka.bDrivesOn := FALSE;                   		 (* Switch on *)
	Kuka.PlcToKuka.bDrivesOff := FALSE;                   		 (* Switch off *)
	tonStatusDelay(IN := FALSE,
				    PT := tStatusDelay);
ELSE

	IF NOT bNoEStop
	     OR NOT bDrivesOn
	THEN
		Kuka.PlcToKuka.bDrivesOn := FALSE;                   		 (* Switch on *)
		Kuka.PlcToKuka.bDrivesOff := FALSE;                   		 (* Switch off *)
	ELSE
		IF Kuka.KukaToPlc.bIOActConf
		     AND NOT Kuka.KukaToPlc.bPeriRdy
		THEN
			Kuka.PlcToKuka.bDrivesOn := TRUE;                   	(* Switch on *)
			Kuka.PlcToKuka.bDrivesOff := TRUE;                   		 (* Switch off *)
		ELSE
			Kuka.PlcToKuka.bDrivesOn := FALSE;                   	 (* Switch on *)
			Kuka.PlcToKuka.bDrivesOff := TRUE;                   		 (* Switch off *)
		END_IF
	END_IF;

END_IF;

Kuka.PlcToKuka.nOverride := LREAL_TO_INT(LIMIT(0,lrOverride,100));

tonStatusDelay(IN := Kuka.KukaToPlc.bPeriRdy,		(* Control enabled *)
			   PT := tStatusDelay);
bStatus := tonStatusDelay.Q;

END_FUNCTION_BLOCK

// ---- POUs/Tc2 Objects/ExternalHardware/KUKA/FB_KUKA_Prg.TcPOU
FUNCTION_BLOCK FB_KUKA_Prg
(*

The function block used to start kuka

Constructor: 		Patryk Panylo
Company:		E. Riexinger GmbH
Date:			18.11.2016
Version:			1.00

Date:			Revision:		Who:				Comment

*)
VAR_INPUT
	(* Input variables / Eingang Variablen *)
	bEnable						:BOOL;			(* Signal FB enable *)
	bReset						:BOOL;			(* Signal reset *)
	bAutoHome					:BOOL;			(* Auto := TRUE, Home := FALSE *)
	bStart						:BOOL;			(* Start program *)
	bStop						:BOOL;			(* Stop program *)
	nProgNo						:INT;			(* Program number *)
	tMaxRefTime					:TIME := t#60s;	(* Maximal referenc time *)
END_VAR
VAR_OUTPUT
	(* Output variables / Ausgang Variablen *)
	bRunning					:BOOL;						(* Program running *)
	bDone						:BOOL;						(* Program done *)
	bBusy						:BOOL;						(* Program busy *)
	bError						:BOOL;						(* Error *)
	udnErrorNo					:UDINT;
END_VAR
VAR_IN_OUT
	(* Input Output variables / Ausgang Variablen *)
	Kuka						:ST_KUKA_REF;
END_VAR
VAR
	(* Enummerations *)
	etKukaStart					:ET_KukaStart;

	(* Variables *)
	bFirstTime					:BOOL;

	nWatchdog					:INT;

	(* References *)

	(* Interfaces *)

	(* Instances *)
	rtStart						:R_TRIG;
	rtStop						:R_TRIG;
	rtReset						:R_TRIG;
	tonWatchdog					:TON;

END_VAR


IF NOT bEnable
THEN
	bDone := FALSE;					(* Program done *)
	bBusy := FALSE;                                  	(* Program not busy *)
	bError := FALSE;                                 	(* Program not error *)
	udnErrorNo := 0;                                 		(* Error number *)

	Kuka.PlcToKuka.bPgReset := FALSE;
	Kuka.PlcToKuka.bExtStart := FALSE;
	Kuka.PlcToKuka.bPgNoParity := FALSE;
	Kuka.PlcToKuka.bPgNoValid := FALSE;

	RETURN;
END_IF;

IF NOT bFirstTime
THEN
	tonWatchdog(IN := FALSE);

	Kuka.PlcToKuka.bPgReset := FALSE;
	Kuka.PlcToKuka.bExtStart := FALSE;
	Kuka.PlcToKuka.bPgNoParity := FALSE;
	Kuka.PlcToKuka.bPgNoValid := FALSE;

	etKukaStart := ET_KukaStart_eWaitExecute;              (* Next step *)

	bFirstTime := TRUE;
END_IF

rtReset(CLK := bReset);

IF rtReset.Q
     AND bError
THEN
	bError := FALSE;

	tonWatchdog(IN := FALSE);

	Kuka.PlcToKuka.bPgReset := FALSE;
	Kuka.PlcToKuka.bExtStart := FALSE;
	Kuka.PlcToKuka.bPgNoParity := FALSE;
	Kuka.PlcToKuka.bPgNoValid := FALSE;

	etKukaStart := ET_KukaStart_eWaitExecute;              (* Next step *)
END_IF

(* Wait for triger *)
rtStart(
	CLK := bStart
);

IF rtStart.Q
     AND Kuka.PlcToKuka.bDrivesOff
     AND Kuka.PlcToKuka.bMoveEnable
     AND Kuka.KukaToPlc.bUserSafe
     AND Kuka.KukaToPlc.bAlarmStop
     AND Kuka.KukaToPlc.bPeriRdy
     AND NOT Kuka.KukaToPlc.bProAct
     AND NOT Kuka.PlcToKuka.bDrivesOn
     AND NOT Kuka.KukaToPlc.bStopMess
THEN
	Kuka.PlcToKuka.bPgReset := FALSE;
	Kuka.PlcToKuka.bExtStart := FALSE;
	Kuka.PlcToKuka.bPgNoParity := FALSE;
	Kuka.PlcToKuka.bPgNoValid := FALSE;
	Kuka.PlcToKuka.nPgNo := 0;

	etKukaStart := ET_KukaStart_eWaitExecute;              (* Next step *)

END_IF

rtStop(
	CLK := bStop
		    OR NOT Kuka.PlcToKuka.bDrivesOff
     		    OR NOT Kuka.PlcToKuka.bMoveEnable
     		    OR NOT Kuka.KukaToPlc.bUserSafe
     		    OR NOT Kuka.KukaToPlc.bAlarmStop
     		    OR NOT Kuka.KukaToPlc.bPeriRdy
     		    OR Kuka.PlcToKuka.bDrivesOn
     		    OR Kuka.KukaToPlc.bStopMess
);

IF rtStop.Q
THEN
	Kuka.PlcToKuka.bPgReset := TRUE;
	Kuka.PlcToKuka.bExtStart := FALSE;
	Kuka.PlcToKuka.bPgNoParity := FALSE;
	Kuka.PlcToKuka.bPgNoValid := FALSE;
	Kuka.PlcToKuka.nPgNo := 0;

	etKukaStart := ET_KukaStart_eWaitExecute;              (* Next step *)

ELSIF NOT Kuka.KukaToPlc.bApplRun
THEN
	Kuka.PlcToKuka.bPgReset := FALSE;
END_IF

bRunning := Kuka.KukaToPlc.bApplRun
		      AND Kuka.KukaToPlc.bProAct;

(* Send command *)
CASE etKukaStart OF

	ET_KukaStart_eWaitExecute:
		bBusy := FALSE;                                     	(* Program not busy *)
		bError := FALSE;                         		(* Program not error *)
		udnErrorNo := 0;                         		(* Error number *)

		IF rtStart.Q
		     AND NOT bStop
		THEN
			nWatchdog := 0;
			bDone:= FALSE;                               		(* Program done *)
			bBusy := TRUE;                                  	(* Program busy *)

			tonWatchdog(IN := FALSE);

			Kuka.PlcToKuka.bExtStart := FALSE;
			Kuka.PlcToKuka.bPgNoParity := FALSE;
			Kuka.PlcToKuka.bPgNoValid := FALSE;
			Kuka.PlcToKuka.nPgNo := nProgNo;

			IF NOT bAutoHome
			     AND Kuka.KukaToPlc.bInHome
			THEN
				etKukaStart := ET_KukaStart_eDone;              (* Next step *)
			ELSE
				etKukaStart := ET_KukaStart_eExtStart;              (* Next step *)
			END_IF

		END_IF

	ET_KukaStart_eExtStart:
		(*nWatchdog := nWatchdog + 1;*)

		Kuka.PlcToKuka.bExtStart := TRUE;
		Kuka.PlcToKuka.bPgNoParity := FALSE;
		Kuka.PlcToKuka.bPgNoValid := FALSE;

		IF Kuka.KukaToPlc.bProAct
		     AND Kuka.KukaToPlc.bOnPath
		     AND NOT Kuka.KukaToPlc.bApplRun
		     AND NOT Kuka.KukaToPlc.bStopMess
		THEN
			nWatchdog := 0;

			(*Kuka.PlcToKuka.bExtStart := FALSE;
			Kuka.PlcToKuka.bPgNoParity := FALSE;
			Kuka.PlcToKuka.bPgNoValid := FALSE;*)

			etKukaStart := ET_KukaStart_eWfInHome;              (* Next step *)

		ELSIF Kuka.KukaToPlc.bStopMess
			    OR nWatchdog > 1000
		THEN
			Kuka.PlcToKuka.bExtStart := FALSE;
			Kuka.PlcToKuka.bPgNoParity := FALSE;
			Kuka.PlcToKuka.bPgNoValid := FALSE;
			
			udnErrorNo := 1;                     (* Error number *)
			
			etKukaStart := ET_KukaStart_eError;              (* Next step *)

		END_IF

	ET_KukaStart_eWfInHome:
		tonWatchdog(
			IN := Kuka.PlcToKuka.nOverride > 0,
			PT:= tMaxRefTime
		);

		IF tonWatchdog.Q
		THEN
			tonWatchdog(IN := FALSE);

			Kuka.PlcToKuka.bExtStart := FALSE;
			Kuka.PlcToKuka.bPgNoParity := FALSE;
			Kuka.PlcToKuka.bPgNoValid := FALSE;

			udnErrorNo := 2;

			etKukaStart := ET_KukaStart_eError;             (* Next step *)

		ELSIF (NOT bAutoHome
			    OR (bAutoHome
				    AND (Kuka.KukaToPlc.bInHome
		     			       OR Kuka.KukaToPlc.arbInHome[1])))
			    AND Kuka.KukaToPlc.bProAct
		    	    AND Kuka.KukaToPlc.bOnPath
			    AND NOT Kuka.KukaToPlc.bApplRun
		     	    AND NOT Kuka.KukaToPlc.bStopMess
		THEN
			tonWatchdog(IN := FALSE);

			(*Kuka.PlcToKuka.bExtStart := FALSE;
			Kuka.PlcToKuka.bPgNoParity := FALSE;
			Kuka.PlcToKuka.bPgNoValid := FALSE;*)

			etKukaStart := ET_KukaStart_eWfPgNoReq;              (* Next step *)

		ELSIF Kuka.KukaToPlc.bStopMess
		THEN
			tonWatchdog(IN := FALSE);

			Kuka.PlcToKuka.bExtStart := FALSE;
			Kuka.PlcToKuka.bPgNoParity := FALSE;
			Kuka.PlcToKuka.bPgNoValid := FALSE;

			udnErrorNo := 3;                     (* Error number *)
			
			etKukaStart := ET_KukaStart_eError;              (* Next step *)

		END_IF

	ET_KukaStart_eWfPgNoReq:
		nWatchdog := nWatchdog + 1;

		IF Kuka.KukaToPlc.bPgNoReq
		     AND Kuka.KukaToPlc.bProAct
		     AND Kuka.KukaToPlc.bOnPath
		     AND NOT Kuka.KukaToPlc.bApplRun
		     AND NOT Kuka.KukaToPlc.bStopMess
		THEN
			(*Kuka.PlcToKuka.bExtStart := FALSE;
			Kuka.PlcToKuka.bPgNoParity := FALSE;
			Kuka.PlcToKuka.bPgNoValid := FALSE;*)

			nWatchdog := 0;

			etKukaStart := ET_KukaStart_ePgNoParity;              (* Next step *)

		ELSIF Kuka.KukaToPlc.bStopMess
			   OR nWatchdog > 1000
		THEN
			Kuka.PlcToKuka.bExtStart := FALSE;
			Kuka.PlcToKuka.bPgNoParity := FALSE;
			Kuka.PlcToKuka.bPgNoValid := FALSE;

			udnErrorNo := 4;                     (* Error number *)
			
			etKukaStart := ET_KukaStart_eError;              (* Next step *)

		END_IF

	ET_KukaStart_ePgNoParity:
		nWatchdog := nWatchdog + 1;

		Kuka.PlcToKuka.bPgNoParity := CHECK_PARITY(in :=  Kuka.PlcToKuka.nPgNo, p := 1);

		IF Kuka.KukaToPlc.bProAct
		     AND Kuka.KukaToPlc.bOnPath
		     AND NOT Kuka.KukaToPlc.bApplRun
		     AND NOT Kuka.KukaToPlc.bStopMess
		THEN
			nWatchdog := 0;

			etKukaStart := ET_KukaStart_ePgNoValid;              (* Next step *)

		ELSIF Kuka.KukaToPlc.bStopMess
			    OR nWatchdog > 1000
		THEN
			Kuka.PlcToKuka.bExtStart := FALSE;
			Kuka.PlcToKuka.bPgNoParity := FALSE;
			Kuka.PlcToKuka.bPgNoValid := FALSE;
			
			udnErrorNo := 5;                     (* Error number *)
			
			etKukaStart := ET_KukaStart_eError;              (* Next step *)

		END_IF

	ET_KukaStart_ePgNoValid:
		Kuka.PlcToKuka.bPgNoValid := TRUE;

		IF NOT Kuka.KukaToPlc.bPgNoReq
		     AND NOT Kuka.KukaToPlc.bInHome
		     AND NOT Kuka.KukaToPlc.arbInHome[1]
		     AND Kuka.KukaToPlc.bProAct
		     AND Kuka.KukaToPlc.bOnPath
		     AND Kuka.KukaToPlc.bApplRun
		     AND NOT Kuka.KukaToPlc.bStopMess
		THEN
			Kuka.PlcToKuka.bExtStart := FALSE;
			Kuka.PlcToKuka.bPgNoParity := FALSE;
			Kuka.PlcToKuka.bPgNoValid := FALSE;

			etKukaStart := ET_KukaStart_eWfProgFinish;              (* Next step *)

		ELSIF Kuka.KukaToPlc.bStopMess
		THEN
			Kuka.PlcToKuka.bExtStart := FALSE;
			Kuka.PlcToKuka.bPgNoParity := FALSE;
			Kuka.PlcToKuka.bPgNoValid := FALSE;

			udnErrorNo := 6;                     (* Error number *)
			
			etKukaStart := ET_KukaStart_eError;              (* Next step *)

		END_IF

	ET_KukaStart_eWfProgFinish:
		IF ((Kuka.KukaToPlc.bInHome
		      AND Kuka.PlcToKuka.nPgNo < 100)
		     OR (Kuka.PlcToKuka.nPgNo >= 100
			    AND Kuka.KukaToPlc.arbInHome[1]))
	     	    AND Kuka.KukaToPlc.bProAct
	    	    AND Kuka.KukaToPlc.bOnPath
		    AND NOT Kuka.KukaToPlc.bApplRun
	     	    AND NOT Kuka.KukaToPlc.bStopMess
		THEN
			Kuka.PlcToKuka.bExtStart := FALSE;
			Kuka.PlcToKuka.bPgNoParity := FALSE;
			Kuka.PlcToKuka.bPgNoValid := FALSE;

			etKukaStart := ET_KukaStart_eDone;              (* Next step *)

		ELSIF Kuka.KukaToPlc.bStopMess
		THEN
			Kuka.PlcToKuka.bExtStart := FALSE;
			Kuka.PlcToKuka.bPgNoParity := FALSE;
			Kuka.PlcToKuka.bPgNoValid := FALSE;

			udnErrorNo := 7;                     (* Error number *)
			
			etKukaStart := ET_KukaStart_eError;              (* Next step *)

		END_IF

	ET_KukaStart_eError:
		bBusy := FALSE;						(* Command busy *)
		bError := TRUE;						(* Command error  *)

		etKukaStart := ET_KukaStart_eNoExecute;

	ET_KukaStart_eDone:
		bDone := TRUE;						(* Command done *)
		bBusy := FALSE;						(* Command busy *)

		etKukaStart := ET_KukaStart_eNoExecute;

	ET_KukaStart_eNoExecute:
		IF NOT bStart
		THEN
			(* Reset outputs *)
			bDone := FALSE;						(* Command done *)
			bBusy := FALSE;						(* Command busy *)
			bError := FALSE;						(* Command error  *)

			nWatchdog := 0;

			Kuka.PlcToKuka.bExtStart := FALSE;
			Kuka.PlcToKuka.bPgNoParity := FALSE;
			Kuka.PlcToKuka.bPgNoValid := FALSE;

			etKukaStart := ET_KukaStart_eWaitExecute;
		END_IF
END_CASE;

END_FUNCTION_BLOCK

// ---- POUs/Tc2 Objects/Logic/Oscat/CHECK_PARITY.TcPOU
FUNCTION CHECK_PARITY : BOOL
(*
CHECK_PARITY checks an input byte IN and an associated paritybit P to
even parity. The output is TRUE if the number of bits in the byte IN have
the value TRUE together with the parity-bit results is an even number.
*)
VAR_INPUT
	in : DWORD;	(* input dword *)
	p : BOOL;	(* Parity-Bit *)
END_VAR


(*
version 1.3	18 feb 2008
programmer 	hugo
tested by	tobias

this function checks for an even partity for a dword and partity bit.

*)

CHECK_PARITY := NOT p;
WHILE in > 0 DO
	CHECK_PARITY := CHECK_PARITY XOR in.0 XOR in.1 XOR in.2 XOR in.3;
	in := SHR(in,4);
END_WHILE;

(* code before rev 1.2
WHILE in > 0 DO
	IF in.0 THEN cnt := cnt + 1; END_IF;
	in := SHR(in,1);
END_WHILE;
check_parity := even(cnt) XOR P;
*)


(* revision history

rev 1.0 HM  1.oct.2006

rev 1.1 hm	10.sep.2007
	changed algorithm to improove performance

rev 1.2	hm	8 dec 2007
	changed algorithm to improove performance

rev 1.3 hm	18. feb 2008
	changed algorithm to improove performance
*)

END_FUNCTION

// ---- POUs/Tc2 Objects/ExternalHardware/KUKA/FB_KUKA_REF.TcPOU
FUNCTION_BLOCK FB_KUKA_REF
VAR_INPUT
	KukaToPlc			:ST_KUKATOPLC;
	PlcToKuka			:ST_PLCTOKUKA;
END_VAR
VAR_OUTPUT

END_VAR
VAR_IN_OUT

END_VAR
VAR

END_VAR

;

END_FUNCTION_BLOCK

// ---- POUs/Tc2 Objects/ExternalHardware/KUKA/FB_KUKA_Reset.TcPOU
FUNCTION_BLOCK FB_KUKA_Reset
(*

The function block used to reset the kuka message.

Constructor: 		Patryk Panylo
Company:		E. Riexinger GmbH
Date:			18.11.2016
Version:			1.00

Date:			Revision:		Who:				Comment

*)
VAR_INPUT
	(* Input variables / Eingang Variablen *)
	bReset						:BOOL;		(* Execut the function block *)
	bExtReset					:BOOL;
END_VAR
VAR_OUTPUT
	(* Output variables / Ausgang Variablen *)
	bDone						:BOOL;			(* Status = TRUE indicates that the axis is ready for operation. *)
	bError						:BOOL;			(* Error *)
	udnErrorNo					:UDINT;			(* Error number *)
	sErrorMsg					:STRING; 		(* Error message *)
END_VAR
VAR_IN_OUT
	(* Input Output variables / Ausgang Variablen *)
	Kuka						:ST_KUKA_REF;
END_VAR
VAR
	(* Enummerations *)

	(* Variables *)

	(* References *)

	(* Interfaces *)

	(* Instances *)
	rtExecute						:R_TRIG;
	rtExtReset					:R_TRIG;
	rtDrivesOk					:R_TRIG;
	tonConfMess					:TON;
END_VAR


rtExecute(CLK := bReset);
rtExtReset(CLK := bExtReset
			       AND Kuka.KukaToPlc.bStopMess);
rtDrivesOk(CLK := Kuka.KukaToPlc.bPeriRdy
	   		        AND Kuka.PlcToKuka.bDrivesOff
			        AND Kuka.KukaToPlc.bStopMess);

tonConfMess(
	IN := Kuka.PlcToKuka.bConfMess,
	PT := t#100ms
);

IF rtExecute.Q
     OR rtExtReset.Q
     OR rtDrivesOk.Q
THEN
	Kuka.PlcToKuka.bConfMess := TRUE;

ELSIF tonConfMess.Q
	   OR NOT Kuka.KukaToPlc.bStopMess
THEN
	Kuka.PlcToKuka.bConfMess := FALSE;
END_IF;
(*
IF NOT Kuka.KukaToPlc.bStopMess       (* Error *)
THEN
	Kuka.PlcToKuka.bConfMess := FALSE;
END_IF;
*)

bDone := bReset
		AND NOT Kuka.KukaToPlc.bStopMess;        (* Error *)

END_FUNCTION_BLOCK

// ---- POUs/Tc2 Objects/ExternalHardware/KUKA/FB_KUKA_StartProg.TcPOU
FUNCTION_BLOCK FB_KUKA_StartProg
(*

The function block used to start kuka

Constructor: 		Patryk Panylo
Company:		E. Riexinger GmbH
Date:			18.11.2016
Version:			1.00

Date:			Revision:		Who:				Comment

*)
VAR_INPUT
	(* Input variables / Eingang Variablen *)
	bEnable						:BOOL;			(* Signal FB enable *)
	bStart						:BOOL;			(* Execute start *)
	nProgNo						:INT;			(* Program number *)
	tMaxRefTime					:TIME := t#60s;	(* Maximal referenc time *)
END_VAR
VAR_OUTPUT
	(* Output variables / Ausgang Variablen *)
	bRunning					:BOOL;						(* Program running *)
	bDone						:BOOL;						(* Program done *)
	bBusy						:BOOL;						(* Program busy *)
	bError						:BOOL;						(* Error *)
	udnErrorNo					:UDINT;
END_VAR
VAR_IN_OUT
	(* Input Output variables / Ausgang Variablen *)
	Kuka						:ST_KUKA_REF;
END_VAR
VAR
	(* Enummerations *)
	etKukaStart					:ET_KukaStart;

	(* Variables *)
	bFirstTime					:BOOL;

	nWatchdog					:INT;

	(* References *)

	(* Interfaces *)

	(* Instances *)
	rtStart						:R_TRIG;
	tonWatchdog					:TON;

END_VAR


IF NOT bEnable
THEN
	bDone := FALSE;					(* Program done *)
	bBusy := FALSE;                                  	(* Program not busy *)
	bError := FALSE;                                 	(* Program not error *)
	udnErrorNo := 0;                                 		(* Error number *)

	Kuka.PlcToKuka.bExtStart := FALSE;
	Kuka.PlcToKuka.bPgNoParity := FALSE;
	Kuka.PlcToKuka.bPgNoValid := FALSE;

	RETURN;
END_IF;

IF NOT bFirstTime
THEN
	tonWatchdog(IN := FALSE);

	Kuka.PlcToKuka.bExtStart := FALSE;
	Kuka.PlcToKuka.bPgNoParity := FALSE;
	Kuka.PlcToKuka.bPgNoValid := FALSE;

	etKukaStart := ET_KukaStart_eWaitExecute;              (* Next step *)

	bFirstTime := TRUE;
END_IF

bRunning := Kuka.KukaToPlc.bApplRun
		      AND Kuka.KukaToPlc.bProAct;

IF NOT Kuka.PlcToKuka.bDrivesOff
     OR NOT Kuka.PlcToKuka.bMoveEnable
     OR NOT Kuka.KukaToPlc.bUserSafe
     OR NOT Kuka.KukaToPlc.bAlarmStop
     OR NOT Kuka.KukaToPlc.bPeriRdy
     OR Kuka.PlcToKuka.bDrivesOn
     OR Kuka.KukaToPlc.bStopMess
THEN
	Kuka.PlcToKuka.bExtStart := FALSE;
	Kuka.PlcToKuka.bPgNoParity := FALSE;
	Kuka.PlcToKuka.bPgNoValid := FALSE;

	etKukaStart := ET_KukaStart_eWaitExecute;              (* Next step *)

	RETURN;
END_IF

(* Wait for triger *)
rtStart(
	CLK := bStart
);

IF rtStart.Q
    AND NOT Kuka.KukaToPlc.bProAct
THEN
	etKukaStart := ET_KukaStart_eWaitExecute;              (* Next step *)

END_IF

(* Send command *)
CASE etKukaStart OF

	ET_KukaStart_eWaitExecute:
		bBusy := FALSE;                                     	(* Program not busy *)
		bError := FALSE;                         		(* Program not error *)
		udnErrorNo := 0;                         		(* Error number *)

		IF rtStart.Q
		THEN
			nWatchdog := 0;
			bDone:= FALSE;                               		(* Program done *)
			bBusy := TRUE;                                  	(* Program busy *)

			tonWatchdog(IN := FALSE);

			Kuka.PlcToKuka.bExtStart := FALSE;
			Kuka.PlcToKuka.bPgNoParity := FALSE;
			Kuka.PlcToKuka.bPgNoValid := FALSE;
			Kuka.PlcToKuka.nPgNo := nProgNo;

			etKukaStart := ET_KukaStart_eExtStart;              (* Next step *)

		END_IF

	ET_KukaStart_eExtStart:
		nWatchdog := nWatchdog + 1;

		Kuka.PlcToKuka.bExtStart := TRUE;
		Kuka.PlcToKuka.bPgNoParity := FALSE;
		Kuka.PlcToKuka.bPgNoValid := FALSE;

		IF Kuka.KukaToPlc.bProAct
		     AND Kuka.KukaToPlc.bOnPath
		     AND NOT Kuka.KukaToPlc.bStopMess
		THEN
			nWatchdog := 0;

			Kuka.PlcToKuka.bExtStart := FALSE;
			Kuka.PlcToKuka.bPgNoParity := FALSE;
			Kuka.PlcToKuka.bPgNoValid := FALSE;

			etKukaStart := ET_KukaStart_eWfInHome;              (* Next step *)

		ELSIF Kuka.KukaToPlc.bStopMess
			    OR nWatchdog > 1000
		THEN
			Kuka.PlcToKuka.bExtStart := FALSE;
			Kuka.PlcToKuka.bPgNoParity := FALSE;
			Kuka.PlcToKuka.bPgNoValid := FALSE;
			
			udnErrorNo := 1;                     (* Error number *)
			
			etKukaStart := ET_KukaStart_eError;              (* Next step *)

		END_IF

	ET_KukaStart_eWfInHome:
		tonWatchdog(
			IN := Kuka.PlcToKuka.nOverride > 0,
			PT:= tMaxRefTime
		);

		IF tonWatchdog.Q
		THEN
			tonWatchdog(IN := FALSE);

			Kuka.PlcToKuka.bExtStart := FALSE;
			Kuka.PlcToKuka.bPgNoParity := FALSE;
			Kuka.PlcToKuka.bPgNoValid := FALSE;

			udnErrorNo := 2;

			etKukaStart := ET_KukaStart_eError;             (* Next step *)

		ELSIF Kuka.KukaToPlc.bInHome
		     	    AND Kuka.KukaToPlc.bProAct
		    	    AND Kuka.KukaToPlc.bOnPath
		     	    AND NOT Kuka.KukaToPlc.bStopMess
		THEN
			tonWatchdog(IN := FALSE);

			Kuka.PlcToKuka.bExtStart := FALSE;
			Kuka.PlcToKuka.bPgNoParity := FALSE;
			Kuka.PlcToKuka.bPgNoValid := FALSE;

			etKukaStart := ET_KukaStart_eWfPgNoReq;              (* Next step *)

		ELSIF Kuka.KukaToPlc.bStopMess
		THEN
			tonWatchdog(IN := FALSE);

			Kuka.PlcToKuka.bExtStart := FALSE;
			Kuka.PlcToKuka.bPgNoParity := FALSE;
			Kuka.PlcToKuka.bPgNoValid := FALSE;

			udnErrorNo := 3;                     (* Error number *)
			
			etKukaStart := ET_KukaStart_eError;              (* Next step *)

		END_IF

	ET_KukaStart_eWfPgNoReq:
		nWatchdog := nWatchdog + 1;

		IF Kuka.KukaToPlc.bPgNoReq
		     AND Kuka.KukaToPlc.bProAct
		     AND Kuka.KukaToPlc.bOnPath
		     AND NOT Kuka.KukaToPlc.bStopMess
		THEN
			Kuka.PlcToKuka.bExtStart := FALSE;
			Kuka.PlcToKuka.bPgNoParity := FALSE;
			Kuka.PlcToKuka.bPgNoValid := FALSE;

			nWatchdog := 0;

			etKukaStart := ET_KukaStart_ePgNoParity;              (* Next step *)

		ELSIF Kuka.KukaToPlc.bStopMess
			   OR nWatchdog > 1000
		THEN
			Kuka.PlcToKuka.bExtStart := FALSE;
			Kuka.PlcToKuka.bPgNoParity := FALSE;
			Kuka.PlcToKuka.bPgNoValid := FALSE;

			udnErrorNo := 4;                     (* Error number *)
			
			etKukaStart := ET_KukaStart_eError;              (* Next step *)

		END_IF

	ET_KukaStart_ePgNoParity:
		nWatchdog := nWatchdog + 1;

		Kuka.PlcToKuka.bPgNoParity := CHECK_PARITY(in :=  Kuka.PlcToKuka.nPgNo, p := 1);

		IF Kuka.KukaToPlc.bProAct
		     AND Kuka.KukaToPlc.bOnPath
		     AND NOT Kuka.KukaToPlc.bStopMess
		THEN
			nWatchdog := 0;

			etKukaStart := ET_KukaStart_ePgNoValid;              (* Next step *)

		ELSIF Kuka.KukaToPlc.bStopMess
			    OR nWatchdog > 1000
		THEN
			Kuka.PlcToKuka.bExtStart := FALSE;
			Kuka.PlcToKuka.bPgNoParity := FALSE;
			Kuka.PlcToKuka.bPgNoValid := FALSE;
			
			udnErrorNo := 5;                     (* Error number *)
			
			etKukaStart := ET_KukaStart_eError;              (* Next step *)

		END_IF

	ET_KukaStart_ePgNoValid:
		Kuka.PlcToKuka.bPgNoValid := TRUE;

		IF NOT Kuka.KukaToPlc.bPgNoReq
		     AND NOT Kuka.KukaToPlc.bInHome
		     AND Kuka.KukaToPlc.bProAct
		     AND Kuka.KukaToPlc.bOnPath
		     AND NOT Kuka.KukaToPlc.bStopMess
		THEN
			Kuka.PlcToKuka.bExtStart := FALSE;
			Kuka.PlcToKuka.bPgNoParity := FALSE;
			Kuka.PlcToKuka.bPgNoValid := FALSE;

			etKukaStart := ET_KukaStart_eWfProgFinish;              (* Next step *)

		ELSIF Kuka.KukaToPlc.bStopMess
		THEN
			Kuka.PlcToKuka.bExtStart := FALSE;
			Kuka.PlcToKuka.bPgNoParity := FALSE;
			Kuka.PlcToKuka.bPgNoValid := FALSE;

			udnErrorNo := 6;                     (* Error number *)
			
			etKukaStart := ET_KukaStart_eError;              (* Next step *)

		END_IF

	ET_KukaStart_eWfProgFinish:
		IF Kuka.KukaToPlc.bInHome
	     	    AND Kuka.KukaToPlc.bProAct
	    	    AND Kuka.KukaToPlc.bOnPath
	     	    AND NOT Kuka.KukaToPlc.bStopMess
		THEN
			Kuka.PlcToKuka.bExtStart := FALSE;
			Kuka.PlcToKuka.bPgNoParity := FALSE;
			Kuka.PlcToKuka.bPgNoValid := FALSE;

			etKukaStart := ET_KukaStart_eDone;              (* Next step *)

		ELSIF Kuka.KukaToPlc.bStopMess
		THEN
			Kuka.PlcToKuka.bExtStart := FALSE;
			Kuka.PlcToKuka.bPgNoParity := FALSE;
			Kuka.PlcToKuka.bPgNoValid := FALSE;

			udnErrorNo := 7;                     (* Error number *)
			
			etKukaStart := ET_KukaStart_eError;              (* Next step *)

		END_IF

	ET_KukaStart_eError:
		bBusy := FALSE;						(* Command busy *)
		bError := TRUE;						(* Command error  *)

		etKukaStart := ET_KukaStart_eNoExecute;

	ET_KukaStart_eDone:
		bDone := TRUE;						(* Command done *)
		bBusy := FALSE;						(* Command busy *)

		etKukaStart := ET_KukaStart_eNoExecute;

	ET_KukaStart_eNoExecute:
		IF NOT bStart
		THEN
			(* Reset outputs *)
			bDone := FALSE;						(* Command done *)
			bBusy := FALSE;						(* Command busy *)
			bError := FALSE;						(* Command error  *)

			nWatchdog := 0;

			Kuka.PlcToKuka.bExtStart := FALSE;
			Kuka.PlcToKuka.bPgNoParity := FALSE;
			Kuka.PlcToKuka.bPgNoValid := FALSE;

			etKukaStart := ET_KukaStart_eWaitExecute;
		END_IF
END_CASE;

END_FUNCTION_BLOCK

// ---- POUs/Tc2 Objects/ExternalHardware/KUKA/FB_MoveToKukaRef.TcPOU
FUNCTION_BLOCK FB_MoveToKukaRef
VAR_INPUT
	stRobotToPlc					:ST_ROBOTTOPLC;
END_VAR
VAR_OUTPUT
	stPlcToRobot					:ST_PLCTOROBOT;
END_VAR
VAR_IN_OUT
	Kuka						:ST_KUKA_REF;				(* The KUKA_REF data type  is an interface between the PLC and the KUKA and contains axis information *)
END_VAR
VAR
	rtForceToBase				:R_TRIG;
	rtForceToWork				:R_TRIG;
	rtCutoffToBase				:R_TRIG;
	rtCutoffToWork				:R_TRIG;

	rtMEStartHeat					:R_TRIG;
	rtMEStopHeat				:R_TRIG;
	rtMEStartExtruding				:R_TRIG;
	rtMEStopExtruding				:R_TRIG;
	rtMEStartFlush				:R_TRIG;
	rtMEStopFlush				:R_TRIG;
END_VAR


(* Set general parameter *)


(* Copy the actual values from the robot to the kuka reference *)
Kuka.KukaToPlc.bPgNoReq := stRobotToPlc.arbyInput[2].0;						(* $OUT[33] - A change of signal requests the higher-level controller to send a program number / PGNO Req-Signalwechsel fordert Leitrechner Programmnr. zu senden *)

Kuka.KukaToPlc.bApplRun := stRobotToPlc.arbyInput[2].1;						(* $OUT[34] - Program is currently being executed / TRUE wenn Programm abgearbeitet wird *)
Kuka.KukaToPlc.bErrToPlc := stRobotToPlc.arbyInput[2].2;						(* $OUT[35] - Error output to PLC / Steuerungs- oder Technologiefehler aufgetreten *)
Kuka.KukaToPlc.bInWorkArea := stRobotToPlc.arbyInput[2].3;					(* $OUT[36] - Robot in work area / Roboter in Bearbeitunsbereich*)

Kuka.KukaToPlc.bIOActConf := stRobotToPlc.arbyInput[0].0;						(* $OUT[140] - This output is TRUE if Automatic External mode is selected and the input $I_O_ACT is TRUE. / *)
Kuka.KukaToPlc.bT1:= stRobotToPlc.arbyInput[0].1;							(* $OUT[993] - Operating mode T1 / Betriebsart T1 *)
Kuka.KukaToPlc.bT2 := stRobotToPlc.arbyInput[0].2;							(* $OUT[994] - Operating mode T2/ Betriebsart T2 *)
Kuka.KukaToPlc.bAut := stRobotToPlc.arbyInput[0].3;							(* $OUT[995] - Operating mode Aut / Betriebsart Aut *)
Kuka.KukaToPlc.bExt := stRobotToPlc.arbyInput[0].4;							(* $OUT[996] - Operating mode Ext / Betriebsart Ext *)
Kuka.KukaToPlc.bOnPath := stRobotToPlc.arbyInput[0].5;						(* $OUT[997] - Set as long as the robot stays on its programmed path / TRUE solange sich Rob. auf programmierten Bahn befindet *)
Kuka.KukaToPlc.bInHome := stRobotToPlc.arbyInput[0].6;						(* $OUT[1000] - Whether or not the robot is in its HOME position  / In Home Position *)
Kuka.KukaToPlc.bStopMess := stRobotToPlc.arbyInput[0].7; 						(* $OUT[1010] - Any message occurring which requires the robot to be stopped / Störung Roboter *)
Kuka.KukaToPlc.bUserSafe := stRobotToPlc.arbyInput[1].0;						(* $OUT[1011] - If the safety fence monitoring switch is opened (AUT mode) or an enabling switch is released (T1 or T2 mode). / Abfrage Schutzgitter(Auto)/Zustimmungsschalter(Test) *)
Kuka.KukaToPlc.bPeriRdy := stRobotToPlc.arbyInput[1].1;						(* $OUT[1012] - Robot drives are switched on / TRUE wenn Roboterantriebe eingeschaltet *)
Kuka.KukaToPlc.bAlarmStop := stRobotToPlc.arbyInput[1].2;						(* $OUT[1013] - Emergency stop / Not Aus *)
Kuka.KukaToPlc.bProAct := stRobotToPlc.arbyInput[1].3;							(* $OUT[1021] - Whenever a process is active / Programmbearbeitung aktiv *)

Kuka.KukaToPlc.arbInHome[1]:= stRobotToPlc.arbyInput[3].1;					(* $OUT[1003] - Whether or not the robot is in its HOME position  / In Home Position *)
Kuka.KukaToPlc.arbInHome[2] := stRobotToPlc.arbyInput[3].2;					(* $OUT[1004] - Whether or not the robot is in its HOME position  / In Home Position *)
Kuka.KukaToPlc.arbInHome[3] := stRobotToPlc.arbyInput[3].3;					(* $OUT[1005] - Whether or not the robot is in its HOME position  / In Home Position *)
Kuka.KukaToPlc.arbInHome[4] := stRobotToPlc.arbyInput[3].4;					(* $OUT[1006] - Whether or not the robot is in its HOME position  / In Home Position *)
Kuka.KukaToPlc.arbInHome[5] := stRobotToPlc.arbyInput[3].5;					(* $OUT[1007] - Whether or not the robot is in its HOME position  / In Home Position *)

rtForceToBase(CLK := stRobotToPlc.arbyInput[12].0); Kuka.KukaToPlc.bForceToBase := rtForceToBase.Q;					(* $OUT[10] - Move force to base position *)
rtForceToWork(CLK := stRobotToPlc.arbyInput[12].1); Kuka.KukaToPlc.bForceToWork := rtForceToWork.Q;					(* $OUT[11] - Move force to work position *)
rtCutoffToBase(CLK := stRobotToPlc.arbyInput[12].2); Kuka.KukaToPlc.bCutoffToBase := rtCutoffToBase.Q;					(* $OUT[12] - Move cutoff to base position *)
rtCutoffToWork(CLK := stRobotToPlc.arbyInput[12].3); Kuka.KukaToPlc.bCutoffToWork := rtCutoffToWork.Q;					(* $OUT[13] - Move cutoffe to work position *)

rtMEStartHeat(CLK := stRobotToPlc.arbyInput[13].0); Kuka.KukaToPlc.bMEStartHeat := rtMEStartHeat.Q;						(* $OUT[18] - Start heat *)
rtMEStopHeat(CLK := stRobotToPlc.arbyInput[13].1); Kuka.KukaToPlc.bMEStopHeat := rtMEStopHeat.Q;						(* $OUT[19] - Stop heat *)
rtMEStartExtruding(CLK := stRobotToPlc.arbyInput[13].2); Kuka.KukaToPlc.bMEStartExtruding := rtMEStartExtruding.Q;			(* $OUT[20] - Start extruding *)
rtMEStopExtruding(CLK := stRobotToPlc.arbyInput[13].3); Kuka.KukaToPlc.bMEStopExtruding := rtMEStopExtruding.Q;			(* $OUT[21] - Stop extruding *)
rtMEStartFlush(CLK := stRobotToPlc.arbyInput[13].4); Kuka.KukaToPlc.bMEStartFlush := rtMEStartFlush.Q;					(* $OUT[22] - Start flush *)
rtMEStopFlush(CLK := stRobotToPlc.arbyInput[13].5); Kuka.KukaToPlc.bMEStopFlush := rtMEStopFlush.Q;					(* $OUT[23] - Stop flush *)
Kuka.KukaToPlc.nMEExtrudingSpeed := BYTE_TO_INT(stRobotToPlc.arbyInput[10]);	(* $OUT[100] - Extruding speed [%] *)

(* Copy the setpoint values from the kuka reference to the robot *)
stPlcToRobot.arbyOutput[4] := INT_TO_BYTE(Kuka.PlcToKuka.nPgNo);		(* $IN[33] - Program number / Programmnummer *)
																	(* $IN[33]  + 8 = $IN[41], PGNO_LENGTH = 8 (max. 16) *)
stPlcToRobot.arbyOutput[2].0 := Kuka.PlcToKuka.bPgNoParity;				(* $IN[41] - Input to which the parity bit is transferred from the higher-level controller / Übertragen des Paritätsbit vom Leitrechner *)
stPlcToRobot.arbyOutput[2].1 := Kuka.PlcToKuka.bPgNoValid;				(* $IN[42] - Input to which the command to read the program number is transferred from the higher-level controller / Einlesen der Programmnumer vom Leitrechener *)

stPlcToRobot.arbyOutput[0].0 := Kuka.PlcToKuka.bDrivesOn;					(* $IN[140] - Switch on the robot drives / Einschalten der Roboterantriebe *)
stPlcToRobot.arbyOutput[0].1 := Kuka.PlcToKuka.bDrivesOff;					(* $IN[141] - Switch off the robot drives / Abschalten der Roboterantriebe *)
stPlcToRobot.arbyOutput[0].2 := Kuka.PlcToKuka.bMoveEnable;				(* $IN[143] - Check the robot drives. TRUE Jogging and program execution are possible / Kontrolle der Roboterantriebe *)
stPlcToRobot.arbyOutput[0].3 := Kuka.PlcToKuka.bIOAct;					(* $IN[1025] - If this input is TRUE, the Automatic External interface is active. Default setting:$IN[1025]. *)
stPlcToRobot.arbyOutput[0].4 := Kuka.PlcToKuka.bConfMess;				(* $IN[142] - Acknowledge error / Quittieren von Fehlermeldungen durch den Leitrechner *)
stPlcToRobot.arbyOutput[0].5 := Kuka.PlcToKuka.bExtStart;					(* $IN[145] - If the I/O interface is active, this input can be set to start or continue a program / Extern Start *)

stPlcToRobot.arbyOutput[0].6 := Kuka.PlcToKuka.bCheckMovena;			(* TRUE MOVE_ENABLE monitoring is activated / Überwachung für MOVE_ENABLE *)

stPlcToRobot.arbyOutput[1].0 := Kuka.PlcToKuka.bPgReset;					(* $IN[148] - Cancel a program / Programm abbrechen *)

stPlcToRobot.arbyOutput[10] := INT_TO_BYTE(Kuka.PlcToKuka.nOverride);	(* $IN[100] - Override *)

stPlcToRobot.arbyOutput[6] := INT_TO_BYTE(Kuka.PlcToKuka.nCutOffDist);						(* $IN[50] - Distance of cutoff *)
stPlcToRobot.arbyOutput[7] := INT_TO_BYTE(SHR(Kuka.PlcToKuka.nCutOffDist,8));

stPlcToRobot.arbyOutput[8] := INT_TO_BYTE(Kuka.PlcToKuka.nExtruderOffDist);					(* $IN[66] - Distance aftre extruder is off *)
stPlcToRobot.arbyOutput[9] := INT_TO_BYTE(SHR(Kuka.PlcToKuka.nExtruderOffDist,8));

stPlcToRobot.arbyOutput[14] := UINT_TO_BYTE(Kuka.PlcToKuka.unExtruderStartTime);				(* $IN[82] - Extruder start time *)
stPlcToRobot.arbyOutput[15] := UINT_TO_BYTE(SHR(Kuka.PlcToKuka.unExtruderStartTime,8));

stPlcToRobot.arbyOutput[12].0 := Kuka.PlcToKuka.bForceInBase;			(* $IN[10] - Force in base position *)
stPlcToRobot.arbyOutput[12].1 := Kuka.PlcToKuka.bForceInWork;			(* $IN[11] - Force in work position *)
stPlcToRobot.arbyOutput[12].2 := Kuka.PlcToKuka.bCutoffInBase;			(* $IN[12] - Cutoff in base position *)
stPlcToRobot.arbyOutput[12].3 := Kuka.PlcToKuka.bCutoffInWork;			(* $IN[13] - Cutoff in work position *)

stPlcToRobot.arbyOutput[13].0 := Kuka.PlcToKuka.bMEHeat;				(* $IN[18] - Heat status ON = TRUE, OFF = FALSE *)
stPlcToRobot.arbyOutput[13].1 := Kuka.PlcToKuka.bMEHeating;			(* $IN[19] - Heating status ON = TRUE, OFF = FALSE *)
stPlcToRobot.arbyOutput[13].2 := Kuka.PlcToKuka.bMEHeated;			(* $IN[20] - Heated status ON = TRUE, OFF = FALSE *)
stPlcToRobot.arbyOutput[13].3 := Kuka.PlcToKuka.bMEExtruding;			(* $IN[21] - Extruder status ON = TRUE, OFF = FALSE *)

END_FUNCTION_BLOCK

// ---- POUs/Tc2 Objects/ExternalHardware/Leister/FB_LeisterExtruder_Extruder.TcPOU
FUNCTION_BLOCK FB_LeisterExtruder_Extruder
(*

The function block used to control heater of Leisetr extruder

Constructor: 		Patryk Panylo
Company:		E. Riexinger GmbH
Date:			09.11.2019
Version:			1.00

Date:			Revision:		Who:				Comment
dd.mm.yyyy		x.xx			Initials			comment

*)
VAR_INPUT
	(* Input variables / Eingang Variablen *)
	bEnable						:BOOL;						(* Enable FB signal *)
	bStart						:BOOL;						(* Start extruder *)
	bStop						:BOOL;						(* Stop extruder *)
	tStartDelay					:TIME := t#0ms;				(* Start delay *)
	tReadyDelay					:TIME := t#0ms;				(* Ready delay *)
	bRelease					:BOOL;						(* Release *)
	nSpeed						:INT;						(* Speed 0 - 100 % *)
	tTimeOut						:TIME := t#10s;				(* Timeout of air ok *)
END_VAR
VAR_OUTPUT
	(* Output variables / Ausgang Variablen *)
	bDone						:BOOL;						(* Program done *)
	bDoneDelay					:BOOL;						(* Program done *)
	bBusy						:BOOL;						(* Program busy *)
	bError						:BOOL;						(* Error *)
	udnErrorNo					:UDINT;
END_VAR
VAR_IN_OUT
	(* Input Output variables / Ausgang Variablen *)
	Leister						:ST_LEISTER_REF;
END_VAR
VAR
	(* Enummerations *)
	etExtruder					:ET_LeisterExtruder;

	(* Variables *)
	nWatchdog					:INT;

	(* References *)

	(* Interfaces *)

	(* Instances *)
	rtStart						:R_TRIG;
	rtStop						:R_TRIG;
	tonStartDelay					:TON;
	tonReadyDelay				:TON;
	tonWatchdog					:TON;
END_VAR


IF NOT bEnable
THEN
	bDone := FALSE;					(* Program done *)
	bBusy := FALSE;                                  	(* Program not busy *)
	bError := FALSE;                                 	(* Program not error *)
	udnErrorNo := 0;                                 		(* Error number *)

	bBusy := bStart OR bStop;
	bDone := bStart OR bStop;
	bDoneDelay := bDone;
	Leister.bRunning := bStart;

	tonWatchdog(IN := FALSE);

	RETURN;
END_IF;

IF NOT Leister.bEnabled
     OR NOT Leister.bReady
     OR NOT Leister.bStartRelease
THEN
	Leister.nExtruderSetSpeed := 0;
ELSE
	Leister.nExtruderSetSpeed := LIMIT(0, nSpeed, 100);
END_IF

(* Wait for triger *)
tonStartDelay(
	IN := bStart,
	PT := tStartDelay
);
rtStart(
	CLK := tonStartDelay.Q
		    AND bRelease
);

rtStop(
	CLK := bStop
);

IF rtStop.Q
THEN
	etExtruder := ET_LeisterExtruder_eWaitExecute;                      						(* Next step *)

END_IF;

tonReadyDelay(
	IN := bDone,
	PT := tReadyDelay
);

bDoneDelay := tonReadyDelay.Q;

CASE etExtruder
OF
	ET_LeisterExtruder_eWaitExecute:
		bBusy := FALSE;                                     	(* Program not busy *)
		bError := FALSE;                         		(* Program not error *)
		udnErrorNo := 0;                         		(* Error number *)

		IF rtStop.Q
		THEN
			nWatchdog := 0;
			bDone := FALSE;                          		(* Program not done *)
			bBusy := TRUE;                                  	(* Program busy *)

			tonWatchdog(IN := FALSE);

			IF Leister.bEnabled
			THEN
				Leister.bStartExtruder := FALSE;
				Leister.bStopExtruder := TRUE;

				etExtruder := ET_LeisterExtruder_eStopExtruder;              (* Next step *)

			ELSE
				udnErrorNo := 1;                     (* Error number *)

				etExtruder :=  ET_LeisterExtruder_eError;             (* Next step *)
			END_IF

		ELSIF rtStart.Q
			    AND bRelease
			    AND nSpeed > 0
			    AND NOT Leister.bLockedInterface
		THEN
			nWatchdog := 0;
			bDone := FALSE;                          		(* Program not done *)
			bBusy := TRUE;                                  	(* Program busy *)

			tonWatchdog(IN := FALSE);

			Leister.bLockedInterface := TRUE;

			IF Leister.bPlastDriveError
			THEN
				Leister.bStartExtruder := FALSE;
				Leister.bStopExtruder := FALSE;

				udnErrorNo := 2;                     (* Error number *)

				etExtruder :=  ET_LeisterExtruder_eError;             (* Next step *)

			ELSIF Leister.bEnabled
			THEN
	  			IF Leister.bReady
			   	     AND Leister.bStartRelease
				THEN
					Leister.bStartExtruder := TRUE;
					Leister.bStopExtruder := FALSE;

					etExtruder := ET_LeisterExtruder_eStartExtruder;              (* Next step *)
				ELSE
					etExtruder := ET_LeisterExtruder_eWfHeaterReady;
				END_IF
			ELSE
				Leister.bStartExtruder := FALSE;
				Leister.bStopExtruder := FALSE;

				udnErrorNo := 3;                     (* Error number *)

				etExtruder :=  ET_LeisterExtruder_eError;             (* Next step *)
			END_IF
		END_IF

	ET_LeisterExtruder_eStartExtruder :
		tonWatchdog(
			IN := TRUE,
			PT:= tTimeOut
		);

		Leister.bStartExtruder := TRUE;
		Leister.bStopExtruder := FALSE;

		IF Leister.bRunning
		THEN
			tonWatchdog(IN := FALSE);

			etExtruder := ET_LeisterExtruder_eDone;             (* Next step *)

		ELSIF Leister.bPlastDriveError
		THEN
			Leister.bStartExtruder := FALSE;
			Leister.bStopExtruder := FALSE;

			tonWatchdog(IN := FALSE);

			udnErrorNo := 4;                     (* Error number *)

			etExtruder := ET_LeisterExtruder_eError;             (* Next step *)

		ELSIF tonWatchdog.Q
		THEN
			Leister.bStartExtruder := FALSE;
			Leister.bStopExtruder := FALSE;

			tonWatchdog(IN := FALSE);

			udnErrorNo := 6;                     (* Error number *)

			etExtruder := ET_LeisterExtruder_eError;             (* Next step *)
		END_IF;

	ET_LeisterExtruder_eStopExtruder :
		tonWatchdog(
			IN := TRUE,
			PT:= tTimeOut
		);

		Leister.bStartExtruder := FALSE;
		Leister.bStopExtruder := TRUE;

		IF NOT Leister.bRunning
		THEN
			tonWatchdog(IN := FALSE);

			etExtruder := ET_LeisterExtruder_eDone;             (* Next step *)

		ELSIF Leister.bPlastDriveError
		THEN
			Leister.bStartExtruder := FALSE;
			Leister.bStopExtruder := FALSE;

			tonWatchdog(IN := FALSE);

			udnErrorNo := 5;                     (* Error number *)

			etExtruder := ET_LeisterExtruder_eError;             (* Next step *)

		ELSIF tonWatchdog.Q
		THEN
			Leister.bStartExtruder := FALSE;
			Leister.bStopExtruder := FALSE;

			tonWatchdog(IN := FALSE);

			udnErrorNo := 6;                     (* Error number *)

			etExtruder := ET_LeisterExtruder_eError;             (* Next step *)
		END_IF;

	ET_LeisterExtruder_eWfHeaterReady:
		tonWatchdog(
			IN := TRUE,
			PT:= tTimeOut
		);

 		 IF Leister.bReady
		      AND Leister.bStartRelease
		THEN
			tonWatchdog(IN := FALSE);

			etExtruder := ET_LeisterExtruder_eStartExtruder;              (* Next step *)

		ELSIF tonWatchdog.Q
			    OR Leister.bPlastDriveError
		THEN
			tonWatchdog(IN := FALSE);

			udnErrorNo := 7;                     (* Error number *)

			etExtruder := ET_LeisterExtruder_eError;             (* Next step *)
		END_IF;

	ET_LeisterExtruder_eError:
		bBusy := FALSE;						(* Command busy *)
		bError := TRUE;						(* Command error  *)

		etExtruder := ET_LeisterExtruder_eNoExecute;

	ET_LeisterExtruder_eDone:
		bDone := TRUE;						(* Command done *)
		bBusy := FALSE;						(* Command busy *)

		etExtruder := ET_LeisterExtruder_eNoExecute;

	ET_LeisterExtruder_eNoExecute:
		IF NOT bStart
		     AND NOT bStop
		THEN
			(* Reset outputs *)
			bDone := FALSE;						(* Command done *)
			bBusy := FALSE;						(* Command busy *)
			bError := FALSE;						(* Command error  *)

			nWatchdog := 0;
			Leister.bLockedInterface := FALSE;

			etExtruder := ET_LeisterExtruder_eWaitExecute;
		END_IF
END_CASE;

END_FUNCTION_BLOCK

// ---- POUs/Tc2 Objects/ExternalHardware/Leister/FB_LeisterExtruder_Heater.TcPOU
FUNCTION_BLOCK FB_LeisterExtruder_Heater
(*

The function block used to control heater of Leisetr extruder

Constructor: 		Patryk Panylo
Company:		E. Riexinger GmbH
Date:			09.11.2019
Version:			1.00

Date:			Revision:		Who:				Comment
dd.mm.yyyy		x.xx			Initials			comment

*)
VAR_INPUT
	(* Input variables / Eingang Variablen *)
	bEnable						:BOOL;						(* Enable FB signal *)
	bStart						:BOOL;						(* Start heater *)
	bStop						:BOOL;						(* Stop heater *)
	bRelease					:BOOL;						(* Release *)
	nAirTemp					:INT;						(* Air temperatur *)
	nPlastTemp					:INT;						(* Plast  temperatur *)
	tTimeOut						:TIME := t#10s;				(* Timeout of air ok *)
END_VAR
VAR_OUTPUT
	(* Output variables / Ausgang Variablen *)
	bDone						:BOOL;						(* Program done *)
	bBusy						:BOOL;						(* Program busy *)
	bError						:BOOL;						(* Error *)
	udnErrorNo					:UDINT;
END_VAR
VAR_IN_OUT
	(* Input Output variables / Ausgang Variablen *)
	Leister						:ST_LEISTER_REF;
END_VAR
VAR
	(* Enummerations *)
	etHeater						:ET_LeisterHeater;

	(* Variables *)
	nWatchdog					:INT;

	(* References *)

	(* Interfaces *)

	(* Instances *)
	rtStart						:R_TRIG;
	rtStop						:R_TRIG;
	tonWatchdog					:TON;
END_VAR


IF NOT bEnable
THEN
	bDone := FALSE;					(* Program done *)
	bBusy := FALSE;                                  	(* Program not busy *)
	bError := FALSE;                                 	(* Program not error *)
	udnErrorNo := 0;                                 		(* Error number *)

	bBusy := bStart OR bStop;
	bDone := bStart OR bStop;
	Leister.bHeating:= bStart;

	tonWatchdog(IN := FALSE);

	RETURN;
END_IF;

(* Wait for triger *)
rtStart(
	CLK := bStart
);

rtStop(
	CLK := bStop
		    OR nAirTemp = 0
		    OR nPlastTemp = 0
);

IF rtStop.Q
THEN
	etHeater := ET_LeisterHeater_eWaitExecute;                      						(* Next step *)

END_IF;

CASE etHeater
OF

	ET_LeisterHeater_eWaitExecute:
		bBusy := FALSE;                                     	(* Program not busy *)
		bError := FALSE;                         		(* Program not error *)
		udnErrorNo := 0;                         		(* Error number *)

		IF rtStop.Q
		THEN
			nWatchdog := 0;
			bDone := FALSE;                          		(* Program not done *)
			bBusy := TRUE;                                  	(* Program busy *)

			tonWatchdog(IN := FALSE);

			IF Leister.bEnabled
			THEN
				Leister.bStartHeater := FALSE;
				Leister.bStopHeater := TRUE;
				Leister.bStartExtruder := FALSE;
				Leister.bStopExtruder := TRUE;

				Leister.nExtruderSetSpeed := 0;

				etHeater := ET_LeisterHeater_eStopHeater;              (* Next step *)

			ELSE
				udnErrorNo := 1;                     (* Error number *)

				etHeater :=  ET_LeisterHeater_eError;             (* Next step *)
			END_IF

		ELSIF rtStart.Q
			    AND bRelease
		   	    AND nAirTemp > 0
		    	    AND nPlastTemp > 0
			    AND NOT Leister.bLockedInterface
		THEN
			nWatchdog := 0;
			bDone := FALSE;                          		(* Program not done *)
			bBusy := TRUE;                                  	(* Program busy *)

			tonWatchdog(IN := FALSE);

			Leister.bLockedInterface := TRUE;

			IF Leister.bAirHeaterError
			    OR Leister.bPlastHeaterError
			THEN
				Leister.bStartHeater := FALSE;
				Leister.bStopHeater := FALSE;
				Leister.bStartExtruder := FALSE;
				Leister.bStopExtruder := FALSE;

				udnErrorNo := 2;                     (* Error number *)

				etHeater :=  ET_LeisterHeater_eError;             (* Next step *)

			ELSIF Leister.bEnabled
			THEN
				Leister.bStartHeater := TRUE;
				Leister.bStopHeater := FALSE;
				Leister.nAirSetTemp := nAirTemp;
				Leister.nPlastSetTemp := nPlastTemp;

				IF Leister.bReady
				     AND Leister.bStartRelease
				THEN
					etHeater := ET_LeisterHeater_eDone;              (* Next step *)
				ELSE
					etHeater := ET_LeisterHeater_eStartHeater;              (* Next step *)
				END_IF
			ELSE
				Leister.bStartHeater := FALSE;
				Leister.bStopHeater := FALSE;
				Leister.bStartExtruder := FALSE;
				Leister.bStopExtruder := FALSE;

				udnErrorNo := 3;                     (* Error number *)

				etHeater :=  ET_LeisterHeater_eError;             (* Next step *)
			END_IF
		END_IF

	ET_LeisterHeater_eStartHeater :
		tonWatchdog(
			IN := TRUE,
			PT:= tTimeOut
		);

		Leister.bStartHeater := TRUE;
		Leister.bStopHeater := FALSE;

		IF Leister.bHeating
		THEN
			tonWatchdog(IN := FALSE);

			etHeater := ET_LeisterHeater_eDone;             (* Next step *)

		ELSIF Leister.bAirHeaterError
		THEN
			Leister.bStartHeater := FALSE;
			Leister.bStopHeater := FALSE;
			Leister.bStartExtruder := FALSE;
			Leister.bStopExtruder := FALSE;;

			tonWatchdog(IN := FALSE);

			udnErrorNo := 4;                     (* Error number *)

			etHeater := ET_LeisterHeater_eError;             (* Next step *)

		ELSIF Leister.bPlastHeaterError
		THEN
			Leister.bStartHeater := FALSE;
			Leister.bStopHeater := FALSE;
			Leister.bStartExtruder := FALSE;
			Leister.bStopExtruder := FALSE;

			tonWatchdog(IN := FALSE);

			udnErrorNo := 5;                     (* Error number *)

			etHeater := ET_LeisterHeater_eError;             (* Next step *)

		ELSIF tonWatchdog.Q
		THEN
			Leister.bStartHeater := FALSE;
			Leister.bStopHeater := FALSE;
			Leister.bStartExtruder := FALSE;
			Leister.bStopExtruder := FALSE;

			tonWatchdog(IN := FALSE);

			udnErrorNo := 6;                     (* Error number *)

			etHeater := ET_LeisterHeater_eError;             (* Next step *)
		END_IF;

	ET_LeisterHeater_eStopHeater :
		tonWatchdog(
			IN := TRUE,
			PT:= tTimeOut
		);

		Leister.bStartHeater := FALSE;
		Leister.bStopHeater := TRUE;
		Leister.bStartExtruder := FALSE;
		Leister.bStopExtruder := TRUE;

		Leister.nExtruderSetSpeed := 0;
		Leister.nAirSetTemp := 0;
		Leister.nPlastSetTemp := 0;

		IF NOT Leister.bHeating
		    AND NOT Leister.bRunning
		    AND NOT Leister.bReady
		    AND NOT Leister.bStartRelease
		THEN
			tonWatchdog(IN := FALSE);

			etHeater := ET_LeisterHeater_eDone;             (* Next step *)

		ELSIF Leister.bAirHeaterError
		THEN
			Leister.bStartHeater := FALSE;
			Leister.bStopHeater := FALSE;
			Leister.bStartExtruder := FALSE;
			Leister.bStopExtruder := FALSE;;

			tonWatchdog(IN := FALSE);

			udnErrorNo := 4;                     (* Error number *)

			etHeater := ET_LeisterHeater_eError;             (* Next step *)

		ELSIF Leister.bPlastHeaterError
		THEN
			Leister.bStartHeater := FALSE;
			Leister.bStopHeater := FALSE;
			Leister.bStartExtruder := FALSE;
			Leister.bStopExtruder := FALSE;

			tonWatchdog(IN := FALSE);

			udnErrorNo := 5;                     (* Error number *)

			etHeater := ET_LeisterHeater_eError;             (* Next step *)

		ELSIF tonWatchdog.Q
		THEN
			Leister.bStartHeater := FALSE;
			Leister.bStopHeater := FALSE;
			Leister.bStartExtruder := FALSE;
			Leister.bStopExtruder := FALSE;

			tonWatchdog(IN := FALSE);

			udnErrorNo := 6;                     (* Error number *)

			etHeater := ET_LeisterHeater_eError;             (* Next step *)
		END_IF;

	ET_LeisterHeater_eError:
		bBusy := FALSE;						(* Command busy *)
		bError := TRUE;						(* Command error  *)

		etHeater := ET_LeisterHeater_eNoExecute;

	ET_LeisterHeater_eDone:
		bDone := TRUE;						(* Command done *)
		bBusy := FALSE;						(* Command busy *)

		etHeater := ET_LeisterHeater_eNoExecute;

	ET_LeisterHeater_eNoExecute:
		IF NOT bStart
		     AND NOT bStop
		THEN
			(* Reset outputs *)
			bDone := FALSE;						(* Command done *)
			bBusy := FALSE;						(* Command busy *)
			bError := FALSE;						(* Command error  *)

			nWatchdog := 0;
			Leister.bLockedInterface := FALSE;

			etHeater := ET_LeisterHeater_eWaitExecute;
		END_IF
END_CASE;

END_FUNCTION_BLOCK

// ---- POUs/Tc2 Objects/ExternalHardware/Leister/FB_LEISTER_EXTRUDER_REF.TcPOU
FUNCTION_BLOCK FB_LEISTER_EXTRUDER_REF
VAR_INPUT
	bEnable						:BOOL;						(* Enable *)
	bResetAlarm					:BOOL;						(* Reset alarm *)
	bDriveAbort					:BOOL;						(* Drive abort *)

	bStartHeater					:BOOL;						(* Heater start *)
	bStopHeater					:BOOL;						(* Heater stop *)
	bStartExtruder				:BOOL;						(* Extruder start *)
	bStopExtruder				:BOOL;						(* Extruder start *)

	bEnabled					:BOOL;						(* Enabled *)
	bError						:BOOL;						(* Error *)
	bAirPressureOk				 :BOOL;						(* Air pressure Ok *)

	bReady						:BOOL;						(* Ready *)
	bHeating						:BOOL;						(* Heating *)
	bStartRelease				:BOOL;						(* Start release *)
	bRunning					:BOOL;						(* Running *)

	bAirHeaterError				:BOOL;						(* Air heater error *)
	bPlastHeaterError				:BOOL;						(* Plast heater error *)
	bPlastDriveError				:BOOL;						(* Plast drive error *)

	nExtruderSetSpeed			:INT;						(* Referenc extruding speed 0 - 100 % *)
	nExtruderSpeedMin			:INT;						(* Minimal extruding speed 0 - 600 Upm *)
	nExtruderSpeedMax			:INT;						(* Maximal extruding speed 0 - 600 Upm *)
	nExtrudingActSpeed			:INT;						(* Current extruding speed Upm *)

	nPlastSetTemp				:INT;						(* Referenc plast temperature  °C *)
	nPlastOffsetTemp				:INT;						(* Offset plast temperature  °C *)
	nPlastTempMin				:INT;						(* Minimal plast temperature  °C *)
	nPlastTempMax				:INT;						(* Maximal plast temperature  °C *)
	nPlastActTemp				:INT;						(* Current plast temperature ° C *)

	nAirSetTemp					:INT;						(* Referenc air temperature  °C *)
	nAirOffsetTemp				:INT;						(* Offset air temperature  °C *)
	nAirTempMin					:INT;						(* Minimal air temperature  °C *)
	nAirTempMax				:INT;						(* Maximal air temperature  °C *)
	nAirActTemp					:INT;						(* Current air temperature ° C *)
	nAirActFlow					:INT;						(* Current air flow l/min *)

	bLockedInterface				:BOOL;						(* Interface lock *)

	stTerminalState				AT %I*:ST_TerminalState;
	stLeisterToPlc				AT %I*:ST_LEISTERTOPLC;
	stPlcToLeister				AT %Q*:ST_PLCTOLEISTER;
END_VAR
VAR_OUTPUT

END_VAR
VAR_IN_OUT

END_VAR
VAR

END_VAR

;

END_FUNCTION_BLOCK

// ---- POUs/Tc2 Objects/ExternalHardware/Munsch/FB_MunschExtruder.TcPOU
FUNCTION_BLOCK FB_MunschExtruder
(*

This function block is used to send and recive data's via KL600x to/from Munsch extruder.

KL600x configuration is 	1200 8-N-1

Constructor: 		Patryk Panylo
Company:		E. Riexinger GmbH
Date:			14.09.2016
Version:			1.00

Date:			Revision:		Who:				Comment
dd.mm.yyyy		x.xx			Initials			comment

*)
VAR_INPUT
	(* Input variables / Eingang Variablen *)
	bEnable						:BOOL;					(* Enable FB *)
	sDeviceNetId					:STRING;				(* Fieldbus master NetId *)
	unSlaveAddr 					:UINT;					(* Fixed address of the slave *)
	sDateTime					:STRING;				(* Current date and time *)
	bReset						:BOOL;					(* Reset *)
	bSendExe					:BOOL;					(* Send execute *)
	tSendPeriod					:TIME := t#0s;				(* Send data every period. If tSendPeriod is 0 then th function is not active *)
	stMunschCmd				:ST_MUNSCH_CMD_Data;
	tTimeOut 					:TIME := t#2s;				(* Timout  *)
END_VAR
VAR_OUTPUT
	(* Output variables / Ausgang Variablen *)
	stMunschRes					:ST_MUNSCH_RES_Data;
	bInterfaceReady				:BOOL;				(* Interface ready to use *)
	bInterfaceError				:BOOL;				(* Interface error *)
	bStringReceived				:BOOL;				(* String received *)
END_VAR
VAR_IN_OUT
	(* Input Output variables / Ausgang Variablen *)
	stRXbuffer 					:ComBuffer;
	stTXbuffer					:ComBuffer;
END_VAR
VAR
	(* Enummerations *)

	(* Variables *)
	sSendString					:STRING;
	sReceivedString				:STRING;

	bFirstTime					:BOOL;					(* First PLC cycle *)

	(* References *)

	(* Interfaces *)

	(* Instances *)
	fbKL600x						:FB_KL600xData;

END_VAR
VAR CONSTANT
	bEnableRTSCTS				:BOOL := FALSE;
	udnBaudrate					:UDINT := 1200;
	unDataBits					:UINT := 8;
	sParity						:STRING := 'N';
	unStopBits					:UINT := 1;
	sStringPrefix					:STRING := '$FC';
	sStringSuffix					:STRING := '';
	byEnRTSCTSSubIndex		:BYTE := 16#01;					(* Subindex of object *)
	wEnRTSCTSIndex			:WORD := 16#8000;                 			 (* Index of object *)
	byBaudrateSubIndex			:BYTE := 16#11;					(* Subindex of object *)
	wBaudrateIndex				:WORD := 16#8000;				(* Index of object *)
	byDataFrameSubIndex			:BYTE := 16#15;					(* Subindex of object *)
	wDataFrameIndex				:WORD := 16#8000;                                     (* Index of object *)
END_VAR


IF NOT bEnable							(* Enable FB *)
THEN
	fbKL600x(
		bEnable := FALSE,
		tTimeOut:= tTimeOut,
		sReceivedString := sReceivedString,
		stRXbuffer := stRXbuffer,
		stTXbuffer := stTXbuffer
	);

	bFirstTime := FALSE;					(* First PLC cycle *)
	RETURN;
END_IF

IF NOT bFirstTime
THEN


	bFirstTime := TRUE;
END_IF

IF bReset
     AND bInterfaceError
THEN
	bInterfaceError := FALSE;
END_IF

sSendString := F_MunschCMD(
	stMunschCmd := stMunschCmd
);

fbKL600x(
	bEnable := TRUE,
	sDeviceNetId:= sDeviceNetId,
	unSlaveAddr:= unSlaveAddr,
	sDateTime:= sDateTime,
	bEnableRTSCTS := bEnableRTSCTS,
	udnBaudrate:= udnBaudrate,
	unDataBits:= unDataBits,
	sParity:= sParity,
	unStopBits:= unStopBits,
	sStringPrefix := sStringPrefix,
	sStringSuffix := sStringSuffix,
	bReset := bReset,
	bSendExe:= bSendExe,
	tSendPeriod:= tSendPeriod,
	sSendString:= sSendString,
	byEnRTSCTSSubIndex := byEnRTSCTSSubIndex,
	wEnRTSCTSIndex := wEnRTSCTSIndex,
	byBaudrateSubIndex := byBaudrateSubIndex,
	wBaudrateIndex := wBaudrateIndex,
	byDataFrameSubIndex	 := byDataFrameSubIndex,
	wDataFrameIndex := wDataFrameIndex,
	tTimeOut:= tTimeOut,
	sReceivedString := sReceivedString,
	stRXbuffer := stRXbuffer,
	stTXbuffer := stTXbuffer,
	bKL600xReady => bInterfaceReady,
	bStringReceived => bStringReceived
 );

stMunschRes := F_MunschRES(
	sResponse := sReceivedString
);

IF fbKL600x.arbError[0]
     OR fbKL600x.arbError[1]
     OR fbKL600x.arbError[2]
     OR (bStringReceived AND stMunschRes.etResponse = ET_MUNSCH_RES_CMDERROR)
THEN
	bInterfaceError := TRUE;
END_IF

END_FUNCTION_BLOCK

// ---- POUs/Tc2 Objects/ExternalHardware/Munsch/F_MunschCMD.TcPOU
FUNCTION F_MunschCMD : STRING							(* Command to Munsch extruder *)
VAR_INPUT
	stMunschCmd			:ST_MUNSCH_CMD_Data;
END_VAR
VAR
	usnBaseMaterialTemp		:USINT := 160;					(* Base material temperature 160 °C *)
	usnBaseAirTemp			:USINT := 160;					(* Base air temperature 160 °C *)
END_VAR


CASE stMunschCmd.etCommand OF

	ET_MUNSCH_CMD_NOCMD:						F_MunschCMD := 'NoCmd';
	ET_MUNSCH_CMD_STARTHEAT:					F_MunschCMD := 'H1';
	ET_MUNSCH_CMD_STOPHEAT:					F_MunschCMD := 'H0';
	ET_MUNSCH_CMD_REQHEATSTATUS:			F_MunschCMD := 'h?';
	ET_MUNSCH_CMD_STARTEXTRUDER:			F_MunschCMD := 'R1';
	ET_MUNSCH_CMD_STOPEXTRUDER:				F_MunschCMD := 'R0';
	ET_MUNSCH_CMD_REQEXTRUDERSTATUS:		F_MunschCMD := 'r?';
	ET_MUNSCH_CMD_SETMATERIALTEMP:			F_MunschCMD := CONCAT('M', CHR(INT_TO_BYTE(MIN(MAX(stMunschCmd.nMaterialTemp - usnBaseMaterialTemp, 0), 240))));
	ET_MUNSCH_CMD_REQMATERIALREFTEMP:		F_MunschCMD := 'm?';
	ET_MUNSCH_CMD_REQMATERIALACTTEMP:		F_MunschCMD := 'n?';
	ET_MUNSCH_CMD_SETAIRTEMP:					F_MunschCMD := CONCAT('A', CHR(INT_TO_BYTE(MIN(MAX(stMunschCmd.nAirTemp - usnBaseAirTemp, 0), 240))));
	ET_MUNSCH_CMD_REQAIRREFTEMP:				F_MunschCMD := 'a?';
	ET_MUNSCH_CMD_REQAIRACTTEMP:				F_MunschCMD := 'b?';
	ET_MUNSCH_CMD_REQSTATUS:					F_MunschCMD := 's?';
ELSE
	F_MunschCMD := 'NoCmd';
END_CASE

END_FUNCTION

// ---- POUs/Tc2 Objects/ExternalHardware/Munsch/F_MunschRES.TcPOU
FUNCTION F_MunschRES : ST_MUNSCH_RES_Data			(* Response from Munsch extruder *)
VAR_INPUT
	sResponse					:STRING	;
END_VAR
VAR
	usnBaseMaterialTemp		:USINT := 160;					(* Base material temperature 160 °C *)
	usnBaseAirTemp			:USINT := 160;					(* Base air temperature 160 °C *)
END_VAR


IF sResponse = 'H1'		THEN	F_MunschRES.etResponse := ET_MUNSCH_RES_STARTHEAT;
ELSIF sResponse = 'H0'	THEN	F_MunschRES.etResponse := ET_MUNSCH_RES_STOPHEAT;
ELSIF sResponse = 'h1'	THEN	F_MunschRES.etResponse := ET_MUNSCH_RES_ACKHEATSTATUSON;
ELSIF sResponse = 'h0'	THEN	F_MunschRES.etResponse := ET_MUNSCH_RES_ACKHEATSTATUSOFF;
ELSIF sResponse = 'R1'	THEN	F_MunschRES.etResponse := ET_MUNSCH_RES_STARTEXTRUDER;
ELSIF sResponse = 'R0'	THEN	F_MunschRES.etResponse := ET_MUNSCH_RES_STOPEXTRUDER;
ELSIF sResponse = 'r1'		THEN	F_MunschRES.etResponse := ET_MUNSCH_RES_ACKEXTRUDERSTATUSON;
ELSIF sResponse = 'r0'		THEN	F_MunschRES.etResponse := ET_MUNSCH_RES_ACKEXTRUDERSTATUSOFF;
ELSIF FIND(sResponse, 'M') = 1		THEN	F_MunschRES.etResponse := ET_MUNSCH_RES_SETMATERIALTEMP; F_MunschRES.nMaterialRefTemp := usnBaseMaterialTemp + ASC(DELETE(sResponse,LEN('M'), FIND(sResponse, 'M')));
ELSIF FIND(sResponse, 'm') = 1 		THEN	F_MunschRES.etResponse := ET_MUNSCH_RES_REQMATERIALREFTEMP; F_MunschRES.nMaterialRefTemp := usnBaseMaterialTemp + ASC(DELETE(sResponse,LEN('m'), FIND(sResponse, 'm')));
ELSIF FIND(sResponse, 'n') = 1 		THEN	F_MunschRES.etResponse := ET_MUNSCH_RES_REQMATERIALACTTEMP; F_MunschRES.nMaterialActTemp := usnBaseMaterialTemp + ASC(DELETE(sResponse,LEN('n'), FIND(sResponse, 'n')));
ELSIF FIND(sResponse, 'A') = 1		THEN	F_MunschRES.etResponse := ET_MUNSCH_RES_SETAIRTEMP; F_MunschRES.nAirRefTemp := usnBaseAirTemp + ASC(DELETE(sResponse,LEN('A'), FIND(sResponse, 'A')));
ELSIF FIND(sResponse, 'a') = 1		THEN	F_MunschRES.etResponse := ET_MUNSCH_RES_REQAIRREFTEMP; F_MunschRES.nAirRefTemp := usnBaseAirTemp + ASC(DELETE(sResponse,LEN('a'), FIND(sResponse, 'a')));
ELSIF FIND(sResponse, 'b') = 1		THEN	F_MunschRES.etResponse := ET_MUNSCH_RES_REQAIRACTTEMP; F_MunschRES.nAirActTemp := usnBaseAirTemp + ASC(DELETE(sResponse,LEN('b'), FIND(sResponse, 'b')));
ELSIF sResponse = 's1'	THEN	F_MunschRES.etResponse := ET_MUNSCH_RES_REQSTATUSHEATED;
ELSIF sResponse = 's0'	THEN	F_MunschRES.etResponse := ET_MUNSCH_RES_REQSTATUSHEATING;
ELSIF sResponse = 'sE'	THEN	F_MunschRES.etResponse := ET_MUNSCH_RES_REQSTATUSERROR;
ELSIF sResponse = 'ER' 	THEN	F_MunschRES.etResponse := ET_MUNSCH_RES_CMDERROR;
ELSE F_MunschRES.etResponse := ET_MUNSCH_RES_NOCMD;
END_IF

END_FUNCTION

// ---- POUs/Tc2 Objects/ExternalHardware/Munsch/FB_MunschExtruderAir.TcPOU
FUNCTION_BLOCK FB_MunschExtruderAir
(*

The function block used to control air pressure.

Constructor: 		Patryk Panylo
Company:		E. Riexinger GmbH
Date:			04.11.2016
Version:			1.00

Date:			Revision:		Who:				Comment
dd.mm.yyyy		x.xx			Initials			comment

*)
VAR_INPUT
	(* Input variables / Eingang Variablen *)
	bEnable					:BOOL;						(* Enable FB signal *)
	bIn						:BOOL;						(* Input signal *)
	bExtruderAirOn			:BOOL;						(* Extruder air on *)
	tAirOk					:TIME := t#5s;					(* Timer to delay output air ok *)
	tAirOff					:TIME := t#5s;					(* Timer to delay output air off *)
	tTimeOut					:TIME := t#5s;					(* Timeout *)
END_VAR
VAR_OUTPUT
	(* Output variables / Ausgang Variablen *)
	bAirOk					:BOOL;						(* Air pressure ok *)
	bAirOn					:BOOL;						(* Air pressure on *)
	bError					:BOOL;						(* Error by no air pressure *)
	udnErrorNo				:UDINT;
	udnMessageNo			:UDINT;
END_VAR
VAR
	(* Enummerations *)

	(* Variables *)

	(* References *)

	(* Interfaces *)

	(* Instances *)
	tonDelayAirOk				:TON;						(* Timer to delay *)
	tofDelayAirOff					:TOF;						(* Timer to delay *)
	fbExtrudingAir					:FB_AirPressure;
END_VAR


IF NOT bEnable
THEN
	fbExtrudingAir(
		bEnable := FALSE
	);

	bAirOk := FALSE;
	RETURN;
END_IF

fbExtrudingAir(
	bEnable := bEnable,
	bIn := bIn,
	bNoEStop := bExtruderAirOn,
	tTimeOut := tTimeOut,
	bError => bError,
	udnErrorNo => udnErrorNo,
	udnMessageNo => udnMessageNo
);

tonDelayAirOk(
	IN := fbExtrudingAir.bOut,
	PT := tAirOk
);

bAirOk := tonDelayAirOk.Q;

tofDelayAirOff(
	IN := fbExtrudingAir.bAirOn,
	PT := tAirOff
);

bAirOn := tofDelayAirOff.Q;

END_FUNCTION_BLOCK

// ---- POUs/Tc2 Objects/ExternalHardware/Munsch/FB_MunschExtruder_AirTemp.TcPOU
FUNCTION_BLOCK FB_MunschExtruder_AirTemp
(*

The function block used to control set material temperature on munschs extruder

Constructor: 		Patryk Panylo
Company:		E. Riexinger GmbH
Date:			18.10.2015
Version:			1.00

Date:			Revision:		Who:				Comment
dd.mm.yyyy		x.xx			Initials			comment

*)
VAR_INPUT
	(* Input variables / Eingang Variablen *)
	bEnable						:BOOL;						(* Enable FB signal *)
	bExecute					:BOOL;						(* Execut the function block *)
	nAirTemp					:INT;						(* Air temperatur *)
	nMinAirTemp					:INT;						(* Minimal air temperatur *)
	nMaxAirTemp				:INT;						(* Maximal air temperatur *)
	nAirTempTolerance			:INT := 5;						(* Air temperatur tolerance*)
END_VAR
VAR_OUTPUT
	(* Output variables / Ausgang Variablen *)
	bAirTempAlarm				:BOOL;						(* Exceeded air temperature tolerance  *)
	bDone						:BOOL;						(* Program done *)
	bBusy						:BOOL;						(* Program busy *)
	bError						:BOOL;						(* Error *)
	udnErrorNo					:UDINT;
END_VAR
VAR_IN_OUT
	(* Input Output variables / Ausgang Variablen *)
	Munsch						:ST_MUNSCH_REF;
END_VAR
VAR
	(* Enummerations *)
	etMunschExtruder				:ET_MunschExtruder;

	(* Variables *)
	nWatchdog					:INT;

	(* References *)

	(* Interfaces *)

	(* Instances *)
	rtExecute						:R_TRIG;

END_VAR

IF NOT bEnable
THEN
	bDone := FALSE;					(* Program done *)
	bBusy := FALSE;                                  	(* Program not busy *)
	bError := FALSE;                                 	(* Program not error *)
	udnErrorNo := 0;                                 		(* Error number *)

	RETURN;
END_IF;

(* Wait for triger *)
rtExecute(CLK := bExecute);

(* Send command *)
CASE etMunschExtruder OF

	ET_MunschExtruder_eWaitExecute:
		IF rtExecute.Q
		THEN
			nWatchdog := 0;

			Munsch.bSetAirTemp := TRUE;
			Munsch.bSetMaterialTemp := FALSE;
			Munsch.bStartHeat := FALSE;
			Munsch.bStopHeat  := FALSE;
			Munsch.bStartExtruding := FALSE;
			Munsch.bStopExtruding  := FALSE;
			Munsch.bReadStatus := FALSE;

			etMunschExtruder := ET_MunschExtruder_eChkInterface;              (* Next step *)
		END_IF

	ET_MunschExtruder_eChkInterface:
		nWatchdog := nWatchdog + 1;

		IF NOT Munsch.bLockedInterface
		THEN
			bBusy := FALSE;                                     	(* Program not busy *)
			bError := FALSE;                         		(* Program not error *)
			udnErrorNo := 0;                         		(* Error number *)

